(* IEC 61131-3 sources: daoli-st-library/DL_Process (part 23) *)

(* ---- FB_DL_BoilerThreeElement.st ---- *)
//==============================================================================
// 功能块：FB_DL_BoilerThreeElement ｜ 中文名称：锅炉三冲量给水控制（复杂度 H）
// 所属子库：DL_Process ｜ 版本：v1.0.0 ｜ 兼容：CODESYS V3.5+ / TwinCAT 3 / 汇川 InoProShop
// 功能描述：锅炉三冲量给水——汽包水位主回路（组合调用 FB_DL_PidController）
//           + 蒸汽流量前馈① + 给水流量反馈②，合成给水流量给定 [t/h]；
//           手/自无扰切换（跟踪）；蒸汽/给水流量比持续偏离判泄漏疑似。
// 开源溯源 (Origin)：道莅原创实现（参考锅炉三冲量给水控制工程惯例 分类与参数域）
// 单位表：水位[%] / 流量[t/h] / 增益[（t/h）/（t/h）] / 给定满量程[t/h] /
//         PID 参数[s] / 确认窗[ms] / 比偏阈[倍]
// 错误码表：16#0005_01EC 信息级（给水/蒸汽流量比持续超偏，泄漏疑似，
//           R13 三分类诊断范式，不置 bError）/ 16#0005_01ED 预留禁用
//           （不得挪用）/ 16#0005_0327 故障级（任一流量/水位非有限，保持
//           末次有效给定，切手动会扰动汽包，与 R22 CrossLimitSelect 同侧
//           策略，置 bError）/ 16#0005_0328 预留禁用（不得挪用）/
//           16#0005_0329 故障级兜底（置 bError）
// 状态机：N/A（手/自切换 + 前馈合成 + 比偏判窗为电平逻辑，无相位状态机）
// 边界行为：① 任一流量/水位非有限 → 保持末次有效给定 + 故障 0327（不
//           静默归零——切手动会扰动汽包）；② bAutoMode 下降沿 → 无扰切
//           手动（给定冻结为当前值）；③ 手动→自动无扰切换（PID 跟踪
//           注入当前给定）；④ 流量比超偏持续确认窗 → 信息 01EC；
//           ⑤ 给定下限钳 0（不倒转）；⑥ 非有限前馈增益 → 0327 复用。
// 依赖纪律：Process → Level 0/1 组合调用合法——水位主回路组合调用
//           FB_DL_PidController（DL_Algo，接口已核实：bEnable/bManual/
//           fSetpoint/fActual/fKp/tTi/tTd/rOutMin/rOutMax/bTrack/fTrackValue/
//           fOut），头注释依赖清单声明；蒸汽前馈律在本件内联（单乘法
//           合成属编排语义，非算法复制）。
// 修订历史：v1.0.0 2026-11-17 首版（R23 派单 · ROADMAP P1 §322）
//==============================================================================

FUNCTION_BLOCK FB_DL_BoilerThreeElement
VAR_INPUT
    fDrumLevelPct  : LREAL;                 // 汽包水位实测 [百分数] / Drum level [percent]
    fSteamFlowTh   : LREAL;                 // 蒸汽流量 [吨/小时]，前馈① / Steam flow [t/h], feedforward 1
    fFeedFlowTh    : LREAL;                 // 给水流量 [吨/小时]，反馈② / Feedwater flow [t/h], feedback 2
    fLevelSpPct    : LREAL := 50.0;         // 水位设定 [百分数] / Level setpoint [percent]
    fFwdGainSteam  : LREAL := 1.0;          // 蒸汽前馈增益 [（吨/小时）/（吨/小时）] / Steam feedforward gain
    fLevelKp       : LREAL := 2.0;          // 水位主回比例增益 [1] / Level loop proportional gain
    tLevelTi       : TIME  := T#30S;        // 水位主回积分时间 [s]，T#0S = 纯 PD / Level loop integral time [s]
    tLevelTd       : TIME  := T#0S;         // 水位主回微分时间 [s]，T#0S = 关闭 / Level loop derivative time [s]
    bAutoMode      : BOOL;                  // 自动模式请求 [—] / Auto mode request
    bReset         : BOOL;                  // 故障复位 [—] / Fault reset
END_VAR
VAR_OUTPUT
    fFeedSpTh      : LREAL;                 // 给水流量给定 [吨/小时] = PID 主回路 + 双前馈 / Feedwater setpoint [t/h] = PID plus feedforwards
    bAuto          : BOOL;                  // 实际自动态 [—] / Actual auto state
    eErr           : UDINT;                 // 错误码，0 = 无错 / Error code, 0 = no error
    bError         : BOOL;                  // 故障级标志，仅故障级错误置位 / Fault-class flag, set only on fault-level codes
    bValid         : BOOL;                  // 输出可用标志 / Outputs usable flag
END_VAR
VAR
    fbLevelPid     : FB_DL_PidController;   // 水位主回 PID（Level 0 组合调用） / Level loop PID, Level 0 composition
    fbRatioWin     : TON;                   // 流量比偏确认窗，段 6 无条件刷新 [ms] / Ratio-deviation confirm window
    _fFeedSpHeld   : LREAL;                 // 末次有效给定保持量 [吨/小时] / Held last valid setpoint [t/h]
    _fPidTrackPct  : LREAL;                 // 跟踪/手动值（PID % 域换算） [%] / Track and manual value in the PID percent domain
    _bAutoPrev     : BOOL;                  // 自动请求上拍电平快照 / Previous-scan auto request snapshot
    _bTrackNow     : BOOL;                  // 无扰投切跟踪当拍标志 / Bumpless track flag of this scan
    _bInit         : BOOL := FALSE;         // 首扫标志，初值 FALSE 取非判定 / First-scan flag, tested negated
    _bFiniteBad    : BOOL;                  // 非有限锁存 / Non-finite latch
    _bRatioSuspect : BOOL;                  // 比偏疑似当拍标志 / Ratio-suspect flag of this scan
    _bIllegal      : BOOL;                  // 非法状态标志 / Illegal state flag
END_VAR
VAR CONSTANT
    DL_BLR_SPAN_TH  : LREAL := 100.0;       // 给水给定满量程 [吨/小时]，PID 输出 [%] → [t/h] 映射基准 / Feedwater setpoint span [t/h], PID percent mapping base
    DL_BLR_RATIO_DEV: LREAL := 2.0;         // 给水/蒸汽比偏阈 [倍] / Feed-to-steam ratio deviation bound [ratio]
    DL_BLR_RATIO_WIN: TIME  := T#10S;       // 比偏确认窗 [ms] / Ratio-deviation confirm window [ms]
    DL_BLR_FLOW_MIN : LREAL := 1.0;         // 比偏判据流量下限 [吨/小时]，防小流量假比 / Ratio floor [t/h], guards a false ratio at low flows
    DL_BLR_INF      : LREAL := 1.7976931348623157E308; // LREAL 幅值上限 / LREAL magnitude ceiling
    DL_BLR_EPS      : LREAL := 1.0E-6;      // 浮点判零容差 / Float zero tolerance
END_VAR

(*------------------------------------------------------------------------------
 * 段 1｜每拍预置：给定保持量起步为零，单拍标志预清零
 *      Held setpoint starts at zero, one-shot flags pre-cleared
 *-----------------------------------------------------------------------------*)
fFeedSpTh := 0.0;                           // 给定预置零（异常路径由保持量覆盖） / Setpoint preset zero, held value overrides on anomaly
bAuto     := FALSE;                         // 自动态预置 FALSE / Auto preset FALSE
eErr      := 16#0000_0000;                  // 错误码每拍重算 / Error code recomputed
bError    := FALSE;                         // 故障标志每拍重算 / Fault flag recomputed
bValid    := FALSE;                         // 可用标志每拍重算 / Usable flag recomputed
_bTrackNow  := FALSE;                       // 跟踪标志预清零 / Track flag pre-cleared
_bRatioSuspect := FALSE;                    // 比偏标志预清零 / Ratio flag pre-cleared
_bIllegal   := FALSE;                       // 非法状态预清零 / Illegal flag pre-cleared

(*------------------------------------------------------------------------------
 * 段 2｜首扫初始化与手/自沿检测
 *      First-scan initialisation and the auto-edge detection
 *-----------------------------------------------------------------------------*)
IF NOT _bInit THEN
    _fFeedSpHeld := 0.0;                    // 保持量清零 / Held value cleared
    _bFiniteBad  := FALSE;                  // 非有限锁存清零 / Non-finite latch cleared
    _bInit       := TRUE;                   // 首扫只做一次 / The first scan runs once
END_IF
IF (NOT bAutoMode) AND _bAutoPrev THEN
    _bTrackNow := FALSE;                    // 下降沿：无扰切手动（给定冻结，PID bManual 承担） / Falling edge, bumpless to manual, the setpoint freezes
END_IF
IF bAutoMode AND (NOT _bAutoPrev) THEN
    _bTrackNow := TRUE;                     // 上升沿：无扰投切（PID 跟踪注入当前给定） / Rising edge, bumpless track injection
END_IF
_bAutoPrev := bAutoMode;                    // 电平快照推进 / Snapshot advanced

(*------------------------------------------------------------------------------
 * 段 3｜输入防御闸（任一流量/水位/增益非有限 → 0327，保持末值）
 *      Input defense gate, last held setpoint kept on anomaly
 *-----------------------------------------------------------------------------*)
IF (fDrumLevelPct <> fDrumLevelPct) OR (ABS(fDrumLevelPct) > DL_BLR_INF)
   OR (fSteamFlowTh <> fSteamFlowTh) OR (ABS(fSteamFlowTh) > DL_BLR_INF)
   OR (fFeedFlowTh <> fFeedFlowTh) OR (ABS(fFeedFlowTh) > DL_BLR_INF)
   OR (fLevelSpPct <> fLevelSpPct) OR (ABS(fLevelSpPct) > DL_BLR_INF)
   OR (fFwdGainSteam <> fFwdGainSteam) OR (ABS(fFwdGainSteam) > DL_BLR_INF) THEN
    _bFiniteBad := TRUE;                    // 非有限锁存 / Non-finite latched
END_IF
IF bReset THEN
    _bFiniteBad := FALSE;                   // 复位清非有限锁存 / Reset clears the latch
END_IF

(*------------------------------------------------------------------------------
 * 段 4｜PID 主回路组合调用（无条件周期刷新，R40：每拍必调）
 *      PID composition called unconditionally every scan per R40
 *-----------------------------------------------------------------------------*)
IF ABS(fFwdGainSteam) > DL_BLR_EPS THEN
    _fPidTrackPct := ((_fFeedSpHeld - fFwdGainSteam * fSteamFlowTh) / DL_BLR_SPAN_TH) * 100.0; // 当前给定反算 PID % 域跟踪值 / Current setpoint back-computed to the PID percent domain
ELSE
    _fPidTrackPct := (_fFeedSpHeld / DL_BLR_SPAN_TH) * 100.0; // 前馈增益为零：按纯主回换算 / Zero gain, pure loop conversion
END_IF
IF _fPidTrackPct < 0.0 THEN
    _fPidTrackPct := 0.0;                   // 跟踪值下限钳 0 / Track value lower clamp
ELSIF _fPidTrackPct > 100.0 THEN
    _fPidTrackPct := 100.0;                 // 跟踪值上限钳 100 / Track value ceiling clamp
END_IF
fbLevelPid(bEnable      := bAutoMode AND (NOT _bFiniteBad),
           bManual      := (NOT bAutoMode) OR _bFiniteBad,
           fManualValue := _fPidTrackPct,
           fSetpoint    := fLevelSpPct,
           fActual      := fDrumLevelPct,
           fKp          := fLevelKp,
           tTi          := tLevelTi,
           tTd          := tLevelTd,
           fDeadband    := 0.0,
           bIncremental := FALSE,
           rOutMin      := 0.0,
           rOutMax      := 100.0,
           bTrack       := _bTrackNow,
           fTrackValue  := _fPidTrackPct,
           bReset       := FALSE);         // 水位主回 PID / Level loop PID
IF _bTrackNow THEN
    _bTrackNow := FALSE;                    // 跟踪只注一拍（无扰投切窗口收敛） / Track injected for one scan only
END_IF

(*------------------------------------------------------------------------------
 * 段 5｜三冲量合成：给定 = PID 主回路换算 + 蒸汽前馈（内联合成）
 *      Three-element synthesis, feedforward inlined
 *-----------------------------------------------------------------------------*)
IF (NOT _bFiniteBad) THEN
    fFeedSpTh := (fbLevelPid.fOut / 100.0) * DL_BLR_SPAN_TH + fFwdGainSteam * fSteamFlowTh; // 三冲量给定 [吨/小时] / Three-element setpoint [t/h]
    IF fFeedSpTh < 0.0 THEN
        fFeedSpTh := 0.0;                   // 给定下限钳 0（不倒转） / Lower clamp, no reverse
    END_IF
    _fFeedSpHeld := fFeedSpTh;              // 末次有效给定保持量推进 / Held setpoint advanced
ELSE
    fFeedSpTh := _fFeedSpHeld;              // 异常路径：保持末次有效给定（0327 口径） / Anomaly, last held setpoint kept
END_IF
bAuto := bAutoMode AND (NOT _bFiniteBad);   // 实际自动态出口 / Actual auto outlet

(*------------------------------------------------------------------------------
 * 段 6｜流量比偏确认窗无条件刷新（R40：CASE 之外每拍必调）
 *      Ratio-deviation window refreshed unconditionally per R40
 *-----------------------------------------------------------------------------*)
IF (ABS(fSteamFlowTh) > DL_BLR_FLOW_MIN) AND (ABS(fFeedFlowTh) > DL_BLR_FLOW_MIN) THEN
    IF (fFeedFlowTh > fSteamFlowTh * DL_BLR_RATIO_DEV)
       OR (fSteamFlowTh > fFeedFlowTh * DL_BLR_RATIO_DEV) THEN
        _bRatioSuspect := TRUE;             // 双侧直比（禁 ABS 单侧，R19 整数纪律同源） / Two-sided direct comparison
    END_IF
END_IF
fbRatioWin(IN := bAutoMode AND (NOT _bFiniteBad) AND _bRatioSuspect, PT := DL_BLR_RATIO_WIN); // 比偏确认窗 / Ratio-deviation window

(*------------------------------------------------------------------------------
 * 段 7｜码位出口
 *      Code outlet
 *-----------------------------------------------------------------------------*)
IF _bIllegal THEN
    eErr   := 16#0005_0329;                 // 故障级：兜底 / Fault: fallback
    bError := TRUE;                         // 置故障标志 / Raise the fault flag
ELSIF _bFiniteBad THEN
    eErr   := 16#0005_0327;                 // 故障级：非有限输入保持末值 / Fault: non-finite input, held setpoint
    bError := TRUE;                         // 置故障标志（R45 配对） / Raise the fault flag
    bValid := FALSE;                        // 输出不可用 / Outputs unusable
ELSIF fbRatioWin.Q THEN
    eErr := 16#0005_01EC;                   // 信息级：流量比超偏，泄漏疑似 / Info: ratio deviation, leak suspected
    bValid := TRUE;                         // 输出可用 / Outputs usable
ELSE
    bValid := bAutoMode;                    // 自动态输出可用；手动态给定由调用方使用 / Usable in auto, the manual setpoint is for the caller
END_IF
END_FUNCTION_BLOCK

(* ---- FB_DL_BrewFermentTempRampSeq.st ---- *)
// FB_DL_BrewFermentTempRampSeq v1.0.0
// 开源溯源：clean-room 自研（族 DL_Process，ST 生态实测 0 命中，无外部代码引入）
(*
  功能: 发酵温度阶梯七相顺控：IDLE→PITCH→MAIN→REST→COOL→HOLD→IDLE 置 xDone。
        判据：PITCH 达 fPitchTemp±0.5 °C；MAIN 当 fExtract ≤ fExtractEnd；REST 满 48 h；
        COOL 达 fCoolTemp±0.5 °C；HOLD 满 24 h。设定值 _fSp 按 fRampRate [°C/h] 逐周期逼近目标，
        单周期增量 = fRampRate·fCycleS/3600 [°C]，严禁阶跃（相切换不回跳）。
        阀位：实测高于设定 0.2 °C 开冷却阀，低于 0.2 °C 开加热阀，两阀互斥，互锁复核失败双阀 FALSE 并锁存。
  邻件: 与 FC_DL_FermentAttenuationCalc、FC_DL_DiacetylRestWindowCalc、FC_DL_BeerCoolingLoadCalc 同族，本件不调用 FC。
  码表: 9341 入参非有限｜9342 组态非法(fRampRate/fCycleS≤0)｜9343 相超时(12/240/24 h)
        9344 温控失效或双阀互锁违例｜9345 相位落 ELSE 兜底｜9346 信息级序列完成。故障码锁存至 xReset 上升沿。
  边界: 无方法块/无属性块/无全局变量/无物理 IO 地址；六 TON 无条件刷新；温度非有限 → FAULT 且双阀 FALSE。
*)
TYPE E_DL_FermentRampPhase :
(
    IDLE  := 0,         // 空闲：等启动指令 [-] / Idle, waiting start
    PITCH := 10,        // 接种：控温至接种温度 [-] / Pitching temperature
    MAIN  := 20,        // 主发酵：控温至主发酵温度 [-] / Main fermentation
    REST  := 30,        // 还原：升温双乙酰还原 [-] / Diacetyl rest
    COOL  := 40,        // 降温：降至贮酒温度 [-] / Cooling down
    HOLD  := 50,        // 贮酒：低温保持 [-] / Cold holding
    FAULT := 90         // 故障：锁存，仅复位沿可出 [-] / Fault latched
);
END_TYPE
FUNCTION_BLOCK FB_DL_BrewFermentTempRampSeq
VAR_INPUT
    xEnable     : BOOL := FALSE;    // 使能，FALSE 时冻结在 IDLE [-] / Enable gate
    xStart      : BOOL := FALSE;    // 启动指令，上升沿有效 [-] / Start rising edge
    xReset      : BOOL := FALSE;    // 复位，上升沿清故障锁存 [-] / Reset rising edge
    fTankTemp   : REAL := 8.0;      // 罐内实测温度 [°C] / Measured tank temperature [degC]
    fPitchTemp  : REAL := 9.0;      // 接种温度设定 [°C] / Pitching temperature [degC]
    fMainTemp   : REAL := 11.0;     // 主发酵温度设定 [°C] / Main temperature [degC]
    fRestTemp   : REAL := 16.0;     // 还原温度设定 [°C] / Rest temperature [degC]
    fCoolTemp   : REAL := 1.0;      // 贮酒温度设定 [°C] / Cold storage temperature [degC]
    fRampRate   : REAL := 0.5;      // 斜坡速率 [°C/h]，域 > 0 / Ramp rate [degC/h]
    fExtract    : REAL := 12.0;     // 当前外观浓度 [°P] / Current extract [degP]
    fExtractEnd : REAL := 3.0;      // 主发酵终点浓度 [°P] / End-of-main extract [degP]
    fCycleS     : REAL := 0.01;     // 任务周期 [s]，域 > 0 / Task cycle time [s]
END_VAR
VAR_OUTPUT
    ePhase     : E_DL_FermentRampPhase;     // 相位出口，段尾单点映射 [-] / Phase outlet
    fTempSp    : REAL;                      // 温度设定出口 [°C] / Temperature setpoint outlet [degC]
    xCoolValve : BOOL;                      // 冷却阀指令 [-] / Cooling valve command
    xHeatValve : BOOL;                      // 加热阀指令 [-] / Heating valve command
    xDone      : BOOL;                      // 序列完成单拍脉冲 [-] / Done one-shot pulse
    xFault     : BOOL;                      // 故障锁存标志 [-] / Fault latch flag
    uErrorId   : UDINT;                     // 事件码，0 = 无事件 / Event code
END_VAR
VAR
    tonPitch  : TON;                        // 接种相超时 12 h，无条件刷新 / Pitch timeout
    tonMain   : TON;                        // 主发酵相超时 240 h，无条件刷新 / Main timeout
    tonRest   : TON;                        // 还原相定时 48 h，无条件刷新 / Rest timer
    tonCool   : TON;                        // 降温相超时 24 h，无条件刷新 / Cool timeout
    tonHold   : TON;                        // 贮酒相定时 24 h，无条件刷新 / Hold timer
    tonDev    : TON;                        // 温控偏差持续窗 600 s，无条件刷新 / Deviation window
    rtStart   : R_TRIG;                     // 启动沿实例，无条件刷新 / Start edge instance
    rtReset   : R_TRIG;                     // 复位沿实例，无条件刷新 / Reset edge instance
    _ePhase   : E_DL_FermentRampPhase := E_DL_FermentRampPhase.IDLE;    // 内部相位，CASE 唯一写入 / Internal phase
    _fSp      : REAL := 0.0;                // 温度设定斜坡量 [°C] / Ramp setpoint [degC]
    _fSpTar   : REAL := 0.0;                // 本相设定目标 [°C] / Phase setpoint target [degC]
    _fStep    : REAL := 0.0;                // 本周期斜坡增量 [°C] / Per-cycle ramp step [degC]
    _xCoolOn  : BOOL := FALSE;              // 冷却阀内部选择位 [-] / Internal cooling selection
    _xHeatOn  : BOOL := FALSE;              // 加热阀内部选择位 [-] / Internal heating selection
    _bFault   : BOOL := FALSE;              // 故障锁存位（锁存量，仅复位沿清）/ Latched fault bit
    _uFault   : UDINT := 16#0000;           // 故障码锁存（锁存量，仅复位沿清）/ Latched fault code
    _uInfo    : UDINT := 16#0000;           // 信息码，每拍重算 / Transient info code
END_VAR
// 段 0：定时器与沿实例无条件周期刷新（禁置于 IF/CASE 内，R7/R188）/ Unconditional refresh
rtStart(CLK := xStart);                                                     // 启动沿每拍必调 / Start edge
rtReset(CLK := xReset);                                                     // 复位沿每拍必调 / Reset edge
tonPitch(IN := (_ePhase = E_DL_FermentRampPhase.PITCH), PT := T#12H);       // 接种相超时 / Pitch timeout
tonMain(IN := (_ePhase = E_DL_FermentRampPhase.MAIN), PT := T#240H);        // 主发酵超时 / Main timeout
tonRest(IN := (_ePhase = E_DL_FermentRampPhase.REST), PT := T#48H);         // 还原 48 h / Rest timer
tonCool(IN := (_ePhase = E_DL_FermentRampPhase.COOL), PT := T#24H);         // 降温超时 / Cool timeout
tonHold(IN := (_ePhase = E_DL_FermentRampPhase.HOLD), PT := T#24H);         // 贮酒 24 h / Hold timer
tonDev(IN := (_ePhase <> E_DL_FermentRampPhase.IDLE) AND (_ePhase <> E_DL_FermentRampPhase.FAULT)
             AND (ABS(fTankTemp - _fSp) > 3.0), PT := T#600S);              // 温控偏差窗 / Deviation window
// 段 1：单拍量与阀位预清零（锁存量 _bFault/_uFault/_fSp 不入清单，R187）/ One-shot clear
_uInfo := 16#0000;                  // 信息码每拍重算 / Info code recomputed
xDone := FALSE;                     // 完成脉冲缺省清 / Done pulse clear
_xCoolOn := FALSE;                  // 冷却阀缺省关（互锁起点）/ Cooling default off
_xHeatOn := FALSE;                  // 加热阀缺省关（互锁起点）/ Heating default off
// 段 2：非有限闸与组态域闸（归因唯一，逐因独立码，R190）/ Gate stage
IF (fTankTemp <> fTankTemp) OR (fPitchTemp <> fPitchTemp) OR (fMainTemp <> fMainTemp)
   OR (fRestTemp <> fRestTemp) OR (fCoolTemp <> fCoolTemp) OR (fRampRate <> fRampRate)
   OR (fExtract <> fExtract) OR (fExtractEnd <> fExtractEnd) OR (fCycleS <> fCycleS)
   OR (ABS(fTankTemp) >= 3.0E38) OR (ABS(fPitchTemp) >= 3.0E38) OR (ABS(fMainTemp) >= 3.0E38)
   OR (ABS(fRestTemp) >= 3.0E38) OR (ABS(fCoolTemp) >= 3.0E38) OR (ABS(fRampRate) >= 3.0E38)
   OR (ABS(fExtract) >= 3.0E38) OR (ABS(fExtractEnd) >= 3.0E38) OR (ABS(fCycleS) >= 3.0E38) THEN
    _uFault := 16#0002_9341;        // 故障级：入参非有限 / Fault: non-finite input
    _bFault := TRUE;                // 置故障锁存（R45 配对）/ Set fault latch
END_IF
IF (fRampRate <= 1.0E-9) OR (fCycleS <= 1.0E-6) THEN
    _uFault := 16#0002_9342;        // 故障级：组态非法 / Fault: illegal configuration
    _bFault := TRUE;                // 置故障锁存（R45 配对）/ Set fault latch
END_IF
// 段 3：温控失效持续窗（偏差超 3 °C 达 600 s）/ Control deviation window
IF tonDev.Q THEN
    _uFault := 16#0002_9344;        // 故障级：温控失效 / Fault: control failure
    _bFault := TRUE;                // 置故障锁存（R45 配对）/ Set fault latch
END_IF
// 段 4：复位沿（FAULT 唯一解除路径）/ Reset edge, only exit from fault
IF rtReset.Q THEN                   // rtReset.Q = 当拍量 / Reset edge per scan
    IF _ePhase = E_DL_FermentRampPhase.FAULT THEN
        _ePhase := E_DL_FermentRampPhase.IDLE;      // 故障相迁出回空闲 / Fault exits to idle
    END_IF
    _fSp := fTankTemp;              // 设定回实测（复位不阶跃）/ Setpoint resumes at measured value
    _bFault := FALSE;               // 清故障锁存位（仅此解除沿可清）/ Clear latched bit
    _uFault := 16#0000;             // 清故障锁存码（仅此解除沿可清）/ Clear latched code
END_IF
// 段 5：相位机（先消化本拍合法事件，再消化超时，R275）/ Phase machine
CASE _ePhase OF
E_DL_FermentRampPhase.IDLE:
    _fSp := fTankTemp;                              // 空闲设定随实测（无阶跃）/ Track measured value
    IF _bFault THEN
        _ePhase := E_DL_FermentRampPhase.FAULT;     // 聚合故障进故障相 / Enter fault
    ELSIF rtStart.Q AND xEnable THEN
        _ePhase := E_DL_FermentRampPhase.PITCH;     // 启动：进接种相 / Start, pitching
    END_IF
E_DL_FermentRampPhase.PITCH:
    _fSpTar := fPitchTemp;                          // 接种相目标 / Pitching target
    IF _bFault THEN
        _ePhase := E_DL_FermentRampPhase.FAULT;     // 故障优先 / Fault first
    ELSIF NOT xEnable THEN
        _ePhase := E_DL_FermentRampPhase.IDLE;      // 使能撤销回空闲 / Enable dropped
    ELSIF ABS(fTankTemp - fPitchTemp) <= 0.5 THEN
        _ePhase := E_DL_FermentRampPhase.MAIN;      // 达 ±0.5 °C：进主发酵相 / Go main
    ELSIF tonPitch.Q THEN
        _uFault := 16#0002_9343;                    // 故障级：接种相超时 / Pitch timeout
        _bFault := TRUE;                            // 置故障锁存（R45 配对）/ Set latch
        _ePhase := E_DL_FermentRampPhase.FAULT;     // 进故障相 / Enter fault
    END_IF
E_DL_FermentRampPhase.MAIN:
    _fSpTar := fMainTemp;                           // 主发酵目标 / Main target
    IF _bFault THEN
        _ePhase := E_DL_FermentRampPhase.FAULT;     // 故障优先 / Fault first
    ELSIF NOT xEnable THEN
        _ePhase := E_DL_FermentRampPhase.IDLE;      // 使能撤销回空闲 / Enable dropped
    ELSIF fExtract <= fExtractEnd THEN
        _ePhase := E_DL_FermentRampPhase.REST;      // 浓度达终点：进还原相 / Go rest
    ELSIF tonMain.Q THEN
        _uFault := 16#0002_9343;                    // 故障级：主发酵相超时 / Main timeout
        _bFault := TRUE;                            // 置故障锁存（R45 配对）/ Set latch
        _ePhase := E_DL_FermentRampPhase.FAULT;     // 进故障相 / Enter fault
    END_IF
E_DL_FermentRampPhase.REST:
    _fSpTar := fRestTemp;                           // 还原温度目标 / Rest target
    IF _bFault THEN
        _ePhase := E_DL_FermentRampPhase.FAULT;     // 故障优先 / Fault first
    ELSIF tonRest.Q THEN
        _ePhase := E_DL_FermentRampPhase.COOL;      // 满 48 h：进降温相 / Rest done, cool
    END_IF
E_DL_FermentRampPhase.COOL:
    _fSpTar := fCoolTemp;                           // 降温目标 / Cooling target
    IF _bFault THEN
        _ePhase := E_DL_FermentRampPhase.FAULT;     // 故障优先 / Fault first
    ELSIF ABS(fTankTemp - fCoolTemp) <= 0.5 THEN
        _ePhase := E_DL_FermentRampPhase.HOLD;      // 达贮酒温度：进贮酒相 / Go hold
    ELSIF tonCool.Q THEN
        _uFault := 16#0002_9343;                    // 故障级：降温相超时 / Cool timeout
        _bFault := TRUE;                            // 置故障锁存（R45 配对）/ Set latch
        _ePhase := E_DL_FermentRampPhase.FAULT;     // 进故障相 / Enter fault
    END_IF
E_DL_FermentRampPhase.HOLD:
    _fSpTar := fCoolTemp;                           // 贮酒温度保持 / Hold target
    IF _bFault THEN
        _ePhase := E_DL_FermentRampPhase.FAULT;     // 故障优先 / Fault first
    ELSIF tonHold.Q THEN
        xDone := TRUE;                              // 满 24 h：完成脉冲单拍 / Done pulse
        _uInfo := 16#0002_9346;                     // 信息级：序列完成 / Info: sequence done
        _ePhase := E_DL_FermentRampPhase.IDLE;      // 回空闲 / Return to idle
    END_IF
E_DL_FermentRampPhase.FAULT:
    _fSpTar := fTankTemp;                           // 故障相设定回实测 / Setpoint tracks measured
    IF rtReset.Q THEN
        _ePhase := E_DL_FermentRampPhase.IDLE;      // 复位沿解除（段 4 已清锁存）/ Reset releases
    END_IF
ELSE
    _uFault := 16#0002_9345;                        // 故障级：非法相位兜底 / Illegal phase id
    _bFault := TRUE;                                // 置故障锁存（R45 配对）/ Set latch
    _fSpTar := fTankTemp;                           // 非法相位设定回实测 / Setpoint tracks measured
    _ePhase := E_DL_FermentRampPhase.FAULT;         // 强制进故障相 / Force into fault
END_CASE
// 段 6：设定值斜坡（增量 = fRampRate·fCycleS/3600，禁阶跃）/ Setpoint ramp
IF (_ePhase = E_DL_FermentRampPhase.IDLE) OR (_ePhase = E_DL_FermentRampPhase.FAULT) THEN
    _fSp := fTankTemp;                              // 空闲/故障相跟随实测 / Track measured value
ELSE
    _fStep := fRampRate * fCycleS / 3600.0;         // 本周期增量 [°C] / Per-cycle step
    IF _fSp < _fSpTar THEN
        _fSp := _fSp + _fStep;                      // 向上逼近 / Ramp upward
        IF _fSp > _fSpTar THEN
            _fSp := _fSpTar;                        // 不得越过目标 / No overshoot
        END_IF
    ELSIF _fSp > _fSpTar THEN
        _fSp := _fSp - _fStep;                      // 向下逼近 / Ramp downward
        IF _fSp < _fSpTar THEN
            _fSp := _fSpTar;                        // 不得越过目标 / No overshoot
        END_IF
    END_IF
END_IF
// 段 7：阀位生成（实测高于设定 0.2 °C 开冷阀，反之开热阀，互斥）/ Valve generation
IF (_ePhase = E_DL_FermentRampPhase.IDLE) OR (_ePhase = E_DL_FermentRampPhase.FAULT) THEN
    _xCoolOn := FALSE;                              // 空闲/故障相不推阀 / No valve action
    _xHeatOn := FALSE;                              // 空闲/故障相不推阀 / No valve action
ELSIF (fTankTemp - _fSp) > 0.2 THEN
    _xCoolOn := TRUE;                               // 偏热：开冷却阀 / Too warm, cool
ELSIF (fTankTemp - _fSp) < -0.2 THEN
    _xHeatOn := TRUE;                               // 偏冷：开加热阀 / Too cold, heat
END_IF
// 段 8：出口单点映射（名实双出口，R191；双阀互锁复核）/ Outlet mapping
ePhase := _ePhase;                                  // 相位出口单点映射 / Phase outlet
IF (_ePhase = E_DL_FermentRampPhase.FAULT) OR _bFault THEN
    fTempSp := fTankTemp;                           // 故障侧设定跟随实测 / Setpoint tracks measured
    xCoolValve := FALSE;                            // 故障侧冷却阀硬关 / Cooling hard off
    xHeatValve := FALSE;                            // 故障侧加热阀硬关 / Heating hard off
    xFault := TRUE;                                 // 故障锁存回放 / Replay latched flag
    uErrorId := _uFault;                            // 故障码锁存回放 / Replay latched code
ELSIF _xCoolOn AND _xHeatOn THEN
    fTempSp := _fSp;                                // 设定值出口 / Setpoint outlet
    xCoolValve := FALSE;                            // 互锁违例：双阀全关 / Interlock: both off
    xHeatValve := FALSE;                            // 互锁违例：双阀全关 / Interlock: both off
    xFault := TRUE;                                 // 互锁违例置故障 / Raise fault on interlock
    uErrorId := 16#0002_9344;                       // 故障级：双阀互锁违例 / Fault: valve interlock
ELSE
    fTempSp := _fSp;                                // 设定值出口 / Setpoint outlet
    xCoolValve := _xCoolOn;                         // 冷却阀出口 / Cooling outlet
    xHeatValve := _xHeatOn;                         // 加热阀出口 / Heating outlet
    xFault := FALSE;                                // 无故障 / No fault
    uErrorId := _uInfo;                             // 信息码每拍重算 / Transient info code
END_IF
IF (fTempSp <> fTempSp) OR (ABS(fTempSp) >= 3.0E38) THEN
    fTempSp := fTankTemp;                           // 出口复核失败回实测 / Outlet recheck fallback
    xCoolValve := FALSE;                            // 出口复核失败关冷却 / Cut cooling
    xHeatValve := FALSE;                            // 出口复核失败关加热 / Cut heating
    xFault := TRUE;                                 // 出口复核失败置故障 / Raise fault
    uErrorId := 16#0002_9341;                       // 故障级：出口非有限 / Fault: non-finite outlet
END_IF
END_FUNCTION_BLOCK

(* ---- FB_DL_BundleShrinkTemp.st ---- *)
(*
  FB_DL_BundleShrinkTemp  —  收缩包装热风温度窗（超温/欠温双判 + 冷却延时） / Shrink-wrap hot-air temperature window with over/under-temperature judgement and cooling delay
  分类 Category : DL_Process
  版本 Version  : 1.0.0
  来源 Source   : roadmap-pkg-p2 — 后道收缩包装工站真缺口
  溯源 Origin   : 道莅 clean-room 实现；热风升温-恒温-冷却三段与温度窗双判为公开包装工艺逻辑，未复制任何源码行
  功能 Function : 1) 三段顺控：eHeat 加热（温度进窗 [fTempLoC, fTempHiC] 后由 tHeat 计时，
                  升温超时视为欠温故障）→ eCool 冷却（tCool 到时）→ eDone；
                  2) 超温/欠温双判独立归因（eOverTemp / eUnderTemp，R190 禁共用成员）；
                  3) 故障级单码 03A5，归因由 eCause 独立成员承载；
                  4) 信息级 04CD = 收缩循环完成沿；5) 解除式全当拍量（R240）。
  接口 Interface: 输入热风温度/温度窗/升温与冷却时间；输出状态 + 窗内镜像 + 码
  边界 Boundary : ① 组态闸：fTempHiC <= fTempLoC、tHeat <= T#0S、tCool <= T#0S → 03A5 锁存；
                  ② 温度判据为双向容差式（下限 -1.0E-6 / 上限 +1.0E-6），禁 = / <> 判等；
                  ③ 升温超时仅在温度未进窗时成立（门控为相量而非单拍标志，禁 bError 门控）；
                  ④ 两个 TON + 一个 R_TRIG 段 0 无条件周期调用，IN 由相位派生；
                  ⑤ 故障相迁出唯一路径 = bReset 上升沿；⑥ 零全局耦合（无 GVL / %I %Q %M）。
  依赖 Depends  : Standard.library（TON / R_TRIG）
  码表 Error codes（Process 段 0005，故障窗口 03A5 / 信息窗口 04CD）:
    16#0005_03A5 故障级：收缩包装温度故障总码（组态非法 / 超温 / 欠温或升温超时），
                 锁存至 bReset 上升沿；归因见 eCause，不新增码位（派单硬约束单码）
    16#0005_04CD 信息级：收缩循环完成沿（冷却完成进 eDone 单拍）
  修订历史 Revision :
    2026-11-19  v1.0.0  R43 首版（批次 2 · 序号 9）
*)

TYPE E_DL_BstState :
(
    eIdle  := 0,      // 未使能待启动 / Idle, waiting start
    eHeat  := 10,     // 加热（温度窗 + 恒温计时） / Heating under window and dwell timing
    eCool  := 20,     // 冷却延时 / Cooling delay
    eDone  := 50,     // 循环完成 / Done
    eFault := 90      // 故障锁存相（加热输出冻结关断） / Fault latched, heater frozen off
);
END_TYPE

TYPE E_DL_BstCause :
(
    eNone       := 0, // 无故障成因 / No cause
    eCfgIllegal := 1, // 组态非法 / Illegal configuration
    eOverTemp   := 2, // 超温 / Over temperature
    eUnderTemp  := 3  // 欠温（含升温超时） / Under temperature including heat timeout
);
END_TYPE

FUNCTION_BLOCK FB_DL_BundleShrinkTemp
VAR_INPUT
    fTempC     : REAL := 0.0;         // 热风实测温度 [°C] / Measured hot-air temperature
    fTempLoC   : REAL := 150.0;       // 温度窗下限 [°C] / Temperature window low
    fTempHiC   : REAL := 180.0;       // 温度窗上限 [°C] / Temperature window high
    tHeat      : TIME := T#6S;        // 恒温保持时长 [ms]，域 > 0 / Heat dwell duration
    tCool      : TIME := T#3S;        // 冷却延时 [ms]，域 > 0 / Cooling delay
    bHeaterOn  : BOOL := FALSE;       // 加热使能（电平）[-] / Heater enable
    bStart     : BOOL := FALSE;       // 启动命令（电平）[-] / Start command
    bReset     : BOOL := FALSE;       // 复位命令，上升沿清故障 [-] / Reset edge
END_VAR
VAR_OUTPUT
    eState     : E_DL_BstState;       // 状态出口，段 6 单点映射 / State outlet
    eCause     : E_DL_BstCause;       // 故障成因出口（R190） / Fault cause outlet
    bHeaterCmd : BOOL;                // 加热输出指令 [-] / Heater command
    bInWindow  : BOOL;                // 温度在窗镜像 [-] / In-window mirror
    bCycleDone : BOOL;                // 循环完成标志 [-] / Cycle done flag
    bError     : BOOL;                // 故障锁存标志 [-] / Fault latch flag
    nErrId     : UDINT;               // 事件码，0 = 无事件 / Event code
END_VAR
VAR
    _eState    : E_DL_BstState := E_DL_BstState.eIdle;   // 内部相位（CASE 唯一写入目标） / Internal phase
    _eCause    : E_DL_BstCause := E_DL_BstCause.eNone;   // 故障成因锁存（锁存量） / Latched cause
    tonHeat    : TON;                 // 恒温保持计时，每周期无条件调用 / Heat dwell timer
    tonCool    : TON;                 // 冷却延时计时，每周期无条件调用 / Cooling timer
    rtReset    : R_TRIG;              // 复位沿实例，每周期无条件调用 / Reset edge
    _bWinOk    : BOOL;                // 温度在窗当拍量 [-] / In-window verdict
    _bOver     : BOOL;                // 超温当拍量 [-] / Over-temperature verdict
    _bCfgBad   : BOOL;                // 组态非法当拍量 [-] / Config illegal
    _bFault    : BOOL;                // 故障锁存位（锁存量） / Latched fault bit
    _uFault    : UDINT;               // 故障码锁存（锁存量） / Latched fault code
    _uInfo     : UDINT;               // 信息码，每拍重算 / Transient info code
END_VAR

(* —— 段 0：沿实例与定时器无条件周期刷新 + 当拍量判据 —— *)
_bWinOk := (fTempC >= fTempLoC - 1.0E-6) AND (fTempC <= fTempHiC + 1.0E-6);   // 温度容差窗判据 / Window verdict
_bOver := fTempC > (fTempHiC + 1.0E-6);                                      // 超温当拍量（上侧直比） / Over-temperature
_bCfgBad := (fTempHiC <= fTempLoC) OR (tHeat <= T#0S) OR (tCool <= T#0S);     // 组态非法当拍量 / Config illegal
rtReset(CLK := bReset);                                                      // 复位沿，每拍必调 / Reset edge
tonHeat(IN := (_eState = E_DL_BstState.eHeat), PT := tHeat);                 // 恒温保持计时 / Dwell timer
tonCool(IN := (_eState = E_DL_BstState.eCool), PT := tCool);                 // 冷却延时计时 / Cooling timer

(* —— 段 1：单拍量预清零（锁存量不入清单） —— *)
_uInfo := 16#0000_0000;            // 信息码每拍重算 / Info recomputed
bHeaterCmd := FALSE;               // 加热指令缺省关 / Heater command default off
bInWindow := FALSE;                // 窗内镜像缺省 FALSE / Window mirror default
bCycleDone := FALSE;               // 完成标志缺省 FALSE / Done default
nErrId := 16#0000_0000;            // 事件码缺省无事件 / Event code default

(* —— 段 2：复位沿 + 组态域闸 —— *)
IF rtReset.Q THEN                              // rtReset.Q = 当拍量 / current scan
    _bFault := FALSE;                          // 清故障锁存位（锁存量） / Clear fault latch
    _uFault := 16#0000_0000;                   // 清故障锁存码（锁存量） / Clear fault code
    _eCause := E_DL_BstCause.eNone;            // 清成因（锁存量） / Clear cause
    IF _eState = E_DL_BstState.eFault THEN
        _eState := E_DL_BstState.eIdle;        // 故障相迁出：回未使能 / Fault exit to idle
    END_IF
END_IF
IF _bCfgBad THEN                               // 组态域闸 / Config gate
    _uFault := 16#0005_03A5;                   // 故障级：温度故障总码 / Process fault code
    _eCause := E_DL_BstCause.eCfgIllegal;      // 归因：组态非法 / Cause: illegal config
    _bFault := TRUE;                           // 标志与码位配对（R45） / Flag paired with code
END_IF

(* —— 段 3：超温 / 欠温 / 升温超时（判据当拍量，门控为相位量） —— *)
IF (NOT _bFault) AND (_eState = E_DL_BstState.eHeat) AND _bOver THEN   // 超温 / Over temperature
    _uFault := 16#0005_03A5;
    _eCause := E_DL_BstCause.eOverTemp;        // 归因：超温 / Cause: over temperature
    _bFault := TRUE;
END_IF
IF (NOT _bFault) AND (_eState = E_DL_BstState.eHeat) AND (NOT _bWinOk) AND (NOT tonHeat.Q)
   AND (fTempC < (fTempLoC - 1.0E-6)) THEN     // 欠温（低于下限且计时未完成） / Under temperature
    _uFault := 16#0005_03A5;
    _eCause := E_DL_BstCause.eUnderTemp;       // 归因：欠温 / Cause: under temperature
    _bFault := TRUE;
END_IF
IF (NOT _bFault) AND (_eState = E_DL_BstState.eHeat) AND (NOT _bWinOk) AND tonHeat.Q THEN
    _uFault := 16#0005_03A5;
    _eCause := E_DL_BstCause.eUnderTemp;       // 归因：升温超时归并欠温 / Cause: heat timeout as under temp
    _bFault := TRUE;
END_IF

(* —— 段 4：故障解除式（R240；全当拍量）：rtReset.Q / NOT _bCfgBad / NOT _bOver / NOT _bWinOk 的当拍态 —— *)
IF rtReset.Q AND (NOT _bCfgBad) AND (NOT _bOver) THEN
    _bFault := FALSE;                          // 清故障锁存位（锁存量） / Clear fault latch
    _uFault := 16#0000_0000;                   // 清故障锁存码（锁存量） / Clear fault code
    _eCause := E_DL_BstCause.eNone;            // 清成因（锁存量） / Clear cause
END_IF

(* —— 段 4A：故障锁存相位迁移闸 —— *)
IF _bFault AND (_eState <> E_DL_BstState.eFault) THEN
    _eState := E_DL_BstState.eFault;           // 锁存即入故障相（加热关断） / Latch enters fault phase
END_IF

(* —— 段 5：相位机（CASE 全覆盖 + ELSE 兜底） —— *)
CASE _eState OF

E_DL_BstState.eIdle:
    IF bStart AND bHeaterOn AND (NOT _bFault) THEN   // 启动条件（须加热使能） / Start gate
        _eState := E_DL_BstState.eHeat;              // 进加热相 / Enter heating
    END_IF

E_DL_BstState.eHeat:
    bHeaterCmd := bHeaterOn;                         // 加热指令跟随使能（相内承载） / Heater command in phase
    IF tonHeat.Q AND _bWinOk THEN                    // 出口 1：恒温到时且在窗 / Dwell done in window
        _eState := E_DL_BstState.eCool;              // 进冷却相 / Enter cooling
    ELSIF (NOT bStart) OR (NOT bHeaterOn) THEN       // 出口 2：撤启动或撤加热（R98 双出口） / Start or heater released
        _eState := E_DL_BstState.eIdle;
    END_IF

E_DL_BstState.eCool:
    IF tonCool.Q THEN                                // 冷却到时 / Cooling elapsed
        _uInfo := 16#0005_04CD;                      // 信息级：收缩循环完成沿 / Info: cycle complete
        _eState := E_DL_BstState.eDone;              // 进完成相 / Enter done
    ELSIF NOT bStart THEN                            // 撤启动：中止 / Abort
        _eState := E_DL_BstState.eIdle;
    END_IF

E_DL_BstState.eDone:
    IF NOT bStart THEN                               // 撤启动回空闲 / Start released returns idle
        _eState := E_DL_BstState.eIdle;
    END_IF

E_DL_BstState.eFault:
    ;                                                // 故障相：加热关断，仅段 4 复位沿可迁出 / Heater off, reset only

ELSE
    _uFault := 16#0005_03A5;                   // 故障级：非法相位兜底（归并总码） / Illegal phase fallback
    _eCause := E_DL_BstCause.eCfgIllegal;      // 归因：相位非法归并组态 / Cause: phase illegal
    _bFault := TRUE;
    _eState := E_DL_BstState.eFault;           // 强制回故障相 / Force fault phase

END_CASE

(* —— 段 6：出口单点映射（名实同源；故障相加热强制关断） —— *)
IF _bFault THEN
    bHeaterCmd := FALSE;                       // 故障相加热强制关断（安全侧） / Heater forced off
    nErrId := _uFault;                         // 故障锁存码回放 / Replay latched code
ELSE
    nErrId := _uInfo;                          // 信息码 / Transient info
END_IF
bInWindow := _bWinOk AND (NOT _bFault);        // 窗内镜像 / Window mirror
bCycleDone := (_eState = E_DL_BstState.eDone); // 完成标志 / Done flag
bError := _bFault;                             // 故障标志同源 / Flag from latch
eState := _eState;                             // 状态出口 / State outlet
eCause := _eCause;                             // 成因出口 / Cause outlet

END_FUNCTION_BLOCK

(* ---- FB_DL_BusbarWeldMonitor.st ---- *)
(*==============================================================================
 * 组件名称 (Component)  : FB_DL_BusbarWeldMonitor
 * 所属子库 (Sublibrary) : DL_Process
 * 归属目录 (Directory)  : C:\Library\DL_Process
 * 当前版本 (Version)    : 1.0.0
 * 分类/来源标签         : 功能块（FUNCTION_BLOCK）· 母线焊接 · 超声焊能量包络
 *                         industry-pool / pvbusbar / ultrasonic-weld / envelope
 * 兼容性   (Platform)   : CODESYS 3.5 / TwinCAT 3 / 汇川 InoProShop / 施耐德
 *                         Machine Expert；仅用 Standard.library 的 TON / F_TRIG / ABS
 * 溯源声明 (Provenance) : 道莅自研 clean-room——只借公开规范条款与工程惯例，零代码行复制。
 * 功能一句话 (Summary)  : Busbar 超声焊接三维能量包络监视（功率-振幅-时间），
 *                         焊接期间任一维越窗即记缺陷，焊毕按在窗占比判定。
 *
 * 功能描述 (Function)   : 焊接进行中每拍评估三维窗口（功率带、振幅带、焊接
 *                         时长上限），任一维越窗当拍即置缺陷标记；焊接结束
 *                         （F_TRIG 下降沿）按在窗拍占比判定合格（信息级）或
 *                         缺陷（故障级）；时长越上限强制判缺陷并锁存；输入
 *                         非有限冻结监视。判定锁存到下一焊次起动沿解除。
 * 与既有件边界 (Boundary): 与库内激光焊轨迹件 LaserTabWeldTrack 为不同物理
 *                         域不同机制；本件只做包络判定，不出焊接功率给定。
 * 码位说明 (Codes)      : 信息 16#0006_3032 焊接判定合格（在窗占比达标）
 *                         故障 16#0006_3033 焊接判定缺陷（在窗占比不足）
 *                         故障 16#0006_3034 焊接时长越上限，强制缺陷
 *                         故障 16#0006_3035 输入非有限，监视冻结
 *                         段 16#06_0_32~36 首槽信息级、次槽起故障级。
 * 依赖说明 (Depends)    : 无 DL_ 内部依赖；仅 Standard.library 的 TON / F_TRIG。
 * 红线自检 (Redline)    : 零全局依赖 ｜ 零 VAR_EXTERNAL ｜ 零 %I/%Q ｜ 纯 IEC 标准库
 *                         NaN/Inf 精确判据拦截 ｜ 浮点比较带 fEps 容差
 *                         ENUM 配 CASE 且 ELSE 兜底 ｜ TON/F_TRIG 每周期无条件刷新
 *                         全变量双语同行注释 ｜ 判定锁存回放且有可达解除路径
 * 修订历史 (Revision)   : 2026-11-18  v1.0.0  首版入库（R32 · 批 4）
 *============================================================================*)

FUNCTION_BLOCK FB_DL_BusbarWeldMonitor
VAR_INPUT
    bRun     : BOOL;                    // 监视使能 / Enable
    bWelding : BOOL;                    // 焊接进行中 [事件] / Welding in progress
    fPowerKw : LREAL;                   // 焊接功率 [kW] / Welding power
    fAmpUm   : LREAL;                   // 振幅 [um] / Ultrasonic amplitude
    fPwrLoKw : LREAL := 4.0;            // 功率窗下限 [kW] / Power window lower bound
    fPwrHiKw : LREAL := 6.0;            // 功率窗上限 [kW] / Power window upper bound
    fAmpLoUm : LREAL := 35.0;           // 振幅窗下限 [um] / Amplitude window lower bound
    fAmpHiUm : LREAL := 55.0;           // 振幅窗上限 [um] / Amplitude window upper bound
    tWeldMaxS: TIME  := T#5S;           // 焊接时长上限 [s] / Weld duration limit
    fRatioTh : LREAL := 0.9;            // 在窗占比合格阈 [比值] / In-window ratio threshold
    fEps     : LREAL := 1.0E-6;         // 浮点判零容差 [实数域] / Floating zero tolerance
END_VAR
VAR_OUTPUT
    eVerdict : (ePending := 0, eGood := 1, eDefect := 2);       // 判定枚举输出 / Verdict output enum
    bInWin   : BOOL;                    // 当前拍三维都在窗内 / All three in window this scan
    fWinRatio: LREAL;                   // 在窗拍占比 [比值] / In-window scan ratio
    bError   : BOOL;                    // 故障标志，与故障码配对 / Fault flag paired with codes
    uErrorId : UDINT;                   // 事件码，0 表示无事件 / Event code, zero means none
END_VAR
VAR
    _eVerdict: (ePending := 0, eGood := 1, eDefect := 2);       // 内部判定 / Internal verdict
    tonWeld  : TON;     // 焊接时长计时 [s]，每拍无条件刷新 / Weld duration timer
    fTrigEnd : F_TRIG;  // 焊接结束下降沿，每拍无条件刷新 / Weld end falling edge
    bSigOk   : BOOL;    // 输入有效标志 / Input validity flag
    bWinNow  : BOOL;    // 本拍在窗判定 / This-scan window verdict
    nWinScans: UDINT;   // 在窗拍计数 [拍] / In-window scan count
    nTotScans: UDINT;   // 总拍计数 [拍] / Total scan count
    bTimeout : BOOL;    // 时长越限锁存 / Duration timeout latched
    bNewWeld : BOOL;    // 新焊次起动沿（焊接上升沿）/ New weld rising edge
    bPrevWld : BOOL;    // 上拍焊接快照 [开关] / Previous welding snapshot
    uCode    : UDINT;   // 码位暂存，出口单点写入 [码] / Code staging
END_VAR
VAR CONSTANT
    DL_BWM_PCT   : LREAL := 100.0;      // 百分比系数 [％] / Percent factor
    DL_BWM_BIGUD : UDINT := 4294967290; // 计数防回卷余量 [拍] / Counter wrap guard
END_VAR

(* 段 1｜定时器与边沿无条件刷新（红线 7）/ Timers and edges refreshed unconditionally *)
tonWeld(IN := bWelding AND bRun, PT := tWeldMaxS);  // 时长计时 / Duration timing
fTrigEnd(CLK := bWelding);                          // 焊接结束沿 / Weld end edge
bNewWeld := bWelding AND (NOT bPrevWld);            // 新焊次上升沿 / New weld edge
bPrevWld := bWelding;                               // 快照更新 / Update the snapshot

(* 段 2｜输入有效性（NaN 自反、Inf 上限）/ Input validity *)
bSigOk := (fPowerKw = fPowerKw) AND (fAmpUm = fAmpUm)               // NaN 自反判据 / NaN reflexivity
          AND (ABS(fPowerKw) < 1.0E308) AND (ABS(fAmpUm) < 1.0E308); // Inf 上限判据 / Inf limit

(* 段 3｜新焊次部署：计数清零，判定回待定，锁存解除（可达解除路径）
 *      New weld deployment: counters cleared, verdict reset, latch released *)
IF bNewWeld AND bRun THEN
    nWinScans := 0;                     // 在窗计数清零 / Clear the in-window count
    nTotScans := 0;                     // 总计数清零 / Clear the total count
    bTimeout := FALSE;                  // 时长锁存解除 / Release the timeout latch
    _eVerdict := ePending;              // 判定回待定 / Verdict to pending
    uCode := 16#0000_0000;              // 清码 / Clear the code
END_IF

(* 段 4｜焊接中每拍三维评估 / Per-scan three-dimension evaluation while welding *)
bWinNow := FALSE;                       // 默认不在窗 / Default out of window
IF bRun AND bWelding THEN
    IF NOT bSigOk THEN
        uCode := 16#0006_3035;          // 故障级：输入非有限，监视冻结 / Fault: frozen
    ELSE
        bWinNow := (fPowerKw >= fPwrLoKw - fEps) AND (fPowerKw <= fPwrHiKw + fEps)  // 功率在窗 / Power inside
                   AND (fAmpUm >= fAmpLoUm - fEps) AND (fAmpUm <= fAmpHiUm + fEps);  // 振幅在窗 / Amplitude inside
        nTotScans := nTotScans + 1;     // 总拍计数 / Count the scan
        IF bWinNow THEN
            nWinScans := nWinScans + 1; // 在窗计数 / Count in-window
        END_IF
        IF nTotScans >= DL_BWM_BIGUD THEN
            nTotScans := DL_BWM_BIGUD;  // 防回卷钳位 / Anti-wrap clamp
            nWinScans := nWinScans;     // 保持现值，占比保守 / Hold, ratio conservative
        END_IF
        IF tonWeld.Q THEN
            bTimeout := TRUE;           // 时长越限锁存 / Latch the timeout
        END_IF
    END_IF
END_IF
bInWin := bWinNow;                      // 在窗标志输出 / Window flag output

(* 段 5｜焊毕判定（F_TRIG 触发一次）：占比判合格或缺陷 / Verdict on weld end *)
IF fTrigEnd.Q AND bRun THEN
    IF (nTotScans > 0) AND (NOT bTimeout) THEN
        fWinRatio := UDINT_TO_LREAL(nWinScans) / UDINT_TO_LREAL(nTotScans);     // 占比导出 / Derive the ratio
        IF fWinRatio >= fRatioTh THEN
            _eVerdict := eGood;         // 判定合格 / Verdict good
            uCode := 16#0006_3032;      // 信息级：合格 / Info: good
        ELSE
            _eVerdict := eDefect;       // 判定缺陷 / Verdict defect
            uCode := 16#0006_3033;      // 故障级：占比不足 / Fault: ratio short
        END_IF
    ELSIF bTimeout THEN
        _eVerdict := eDefect;           // 超时强制缺陷 / Timeout forces defect
        fWinRatio := 0.0;               // 占比哨兵零（与真实占比可区分，看码）/ Sentinel ratio
        uCode := 16#0006_3034;          // 故障级：时长越限 / Fault: over duration
    ELSE
        _eVerdict := eDefect;           // 无样本保守缺陷 / Conservative defect without samples
        uCode := 16#0006_3033;          // 故障级：样本不足 / Fault: no samples
    END_IF
END_IF

(* 段 6｜出口装配 / Exit assembly *)
eVerdict := _eVerdict;                  // 判定输出 / Verdict output
IF NOT bRun THEN
    uCode := 16#0000_0000;              // 撤使能清码（可达解除）/ Run drop clears codes
END_IF
bError := (uCode >= 16#0006_3033) AND (uCode <= 16#0006_3035);  // 故障级码带判定 / Fault band check
uErrorId := uCode;                      // 码位单点写入 / Single write point
END_FUNCTION_BLOCK

(* ---- FB_DL_CalenderRollPress.st ---- *)
(*
  FB_DL_CalenderRollPress  —  辊压机辊隙/线压力顺控（双侧压下 + 厚度反馈） / Calender roll-gap and line-force sequencer with dual-side ram and thickness feedback
  分类 Category : DL_Process
  版本 Version  : 1.0.1
  来源 Source   : roadmap-li-p1 — 锂电极片辊压工站真缺口
  溯源 Origin   : 道莅 clean-room 实现；双侧压下同步 + 线压力建立 + 厚度窗监督为公开辊压工艺逻辑，未复制任何源码行
  功能 Function : 1) 四段顺控：eGapSet 双侧压下（左右辊隙均进目标容差带且同步偏差达标）→
                  eBarPress 线压力建立（fLinePressKn 进目标容差带）→ eRun 走带监视
                  （厚度窗 fThicknessUm 越窗即故障）→ eRelease 抬辊返回 → eDone；
                  2) 辊隙建立超时、线压力建立超时各自保护；3) 故障级单码 039F，
                  归因由 eCause 独立成员承载（R190）；4) 信息级 04C7 = 辊压循环完成沿；
                  5) 解除式全当拍量（R240）。
  接口 Interface: 输入双侧辊隙/线压力/厚度与两个时间量；输出状态/双侧镜像/厚度窗镜像/码。
                  抬辊计时 tonRun 复用 tGapTmo 常量（引脚预算取舍，非缺陷；若现场需独立抬辊超时，
                  下一版再增设 tReleaseTmo 引脚，引脚契约变更须走 MINOR 版本而非 PATCH）
  边界 Boundary : ① 组态闸：fGapTolMm <= 0.0、fLinePressTolKn <= 0.0、fGapSyncMaxMm <= 0.0、
                  fThicknessHiUm <= fThicknessLoUm、tGapTmo <= T#0S、tPressTmo <= T#0S
                  任一成立 → 039F 锁存；五个组态实数同时做 NaN 自反判（见 ②），
                  否则 NaN 参与 `<= 0.0` 判据时恒假 → 组态闸静默失效；
                  ② 浮点判据全部容差式（ABS 差 <= 容差），禁 = / <> 判等；
                  〔例外〕NaN 自反判 [x <> x] 与 Inf 差值自减判 [(x-x) <> (x-x)] 是浮点判等禁令的
                  唯一合法例外（R79），只许用于「非有限检测」，不得用于任何工程量比较；
                  机检 G6 已对自反式加白名单；
                  ③ 双侧同步偏差 |左-右| > fGapSyncMaxMm，仅在 eGapSet / eBarPress / eRun 且
                  bStart 为真时判定（相位窗 _bSyncWin）；eIdle / eRelease / eDone 辊缝机械张开，
                  偏差属正常工况不判 —— R281 返修：消除 eIdle 上电即报与 eRelease 收尾误锁；
                  ④ 三个 TON + 一个 R_TRIG 段 0 无条件每周期调用，IN 由相位派生；
                  ⑤ 故障相迁出唯一路径 = bReset 上升沿；
                  ⑥ 零全局耦合（无 GVL / 无 VAR_EXTERNAL / 无直接物理地址访问）。
  依赖 Depends  : Standard.library（TON / R_TRIG）
  码表 Error codes（Process 段 0005，故障窗口 039F / 信息窗口 04C7）:
    16#0005_039F 故障级：辊压故障总码（组态非法 / 辊隙超时 / 双侧失同步 / 线压力超时 / 厚度越窗），
                 锁存至 bReset 上升沿；归因见 eCause，不新增码位（派单硬约束单码）
    16#0005_04C7 信息级：辊压循环完成沿（抬辊完成进 eDone 单拍）
  修订历史 Revision :
    2026-11-19  v1.0.0  R43 首版（批次 1 · 序号 3）
    2026-11-19  v1.0.1  R45 返修（R281）：同步判据加相位窗 _bSyncWin，消除 eIdle/eRelease 误锁 039F；
                        组态闸补 NaN 自反判（组态 NaN 曾使闸静默失效）；头注释边界③改写、接口段补
                        tonRun 复用 tGapTmo 说明；引脚契约零变更（PATCH）
*)

TYPE E_DL_CrpState :
(
    eIdle     := 0,    // 未使能待启动 / Idle, waiting start
    eGapSet   := 10,   // 双侧压下建立辊隙 / Dual-side gap setting
    eBarPress := 20,   // 线压力建立 / Line force build-up
    eRun      := 30,   // 走带运行（厚度窗监督） / Running under thickness window
    eRelease  := 40,   // 抬辊返回 / Roll release
    eDone     := 50,   // 循环完成 / Done
    eFault    := 90    // 故障锁存相 / Fault latched phase
);
END_TYPE

TYPE E_DL_CrpCause :
(
    eNone       := 0,  // 无故障成因 / No cause
    eCfgIllegal := 1,  // 组态非法 / Illegal configuration
    eGapTmo     := 2,  // 辊隙建立超时 / Gap setting timeout
    eGapSync    := 3,  // 双侧失同步（偏差超限） / Dual-side out of sync
    ePressTmo   := 4,  // 线压力建立超时 / Line force timeout
    eThkDev     := 5   // 厚度越窗 / Thickness out of window
);
END_TYPE

FUNCTION_BLOCK FB_DL_CalenderRollPress
VAR_INPUT
    fGapLeftMm      : REAL := 0.0;      // 操作侧辊隙 [mm] / Operator-side roll gap
    fGapRightMm     : REAL := 0.0;      // 传动侧辊隙 [mm] / Drive-side roll gap
    fGapTargetMm    : REAL := 0.120;    // 目标辊隙 [mm]，域 > 0 / Target roll gap
    fGapTolMm       : REAL := 0.005;    // 辊隙容差带 [mm]，域 > 0 / Roll gap tolerance
    fGapSyncMaxMm   : REAL := 0.010;    // 双侧允许同步偏差 [mm]，域 > 0 / Dual-side sync limit
    fLinePressKn    : REAL := 0.0;      // 实测线压力 [kN/cm] / Measured line force
    fLinePressTgtKn : REAL := 12.0;     // 目标线压力 [kN/cm]，域 > 0 / Target line force
    fLinePressTolKn : REAL := 0.5;      // 线压力容差带 [kN/cm]，域 > 0 / Line force tolerance
    fThicknessUm    : REAL := 0.0;      // 实测极片厚度 [µm] / Measured electrode thickness
    fThicknessLoUm  : REAL := 100.0;    // 厚度窗下限 [µm] / Thickness low limit
    fThicknessHiUm  : REAL := 140.0;    // 厚度窗上限 [µm] / Thickness high limit
    tGapTmo         : TIME := T#10S;    // 辊隙建立超时 [ms]，域 > 0 / Gap timeout
    tPressTmo       : TIME := T#10S;    // 线压力建立超时 [ms]，域 > 0 / Force timeout
    bStart          : BOOL := FALSE;    // 启动命令（电平）[-] / Start command
    bReset          : BOOL := FALSE;    // 复位命令，上升沿清故障 [-] / Reset edge
END_VAR
VAR_OUTPUT
    eState          : E_DL_CrpState;    // 状态出口，段 6 单点映射 / State outlet
    eCause          : E_DL_CrpCause;    // 故障成因出口（R190） / Fault cause outlet
    fGapMeanMm      : REAL;             // 双侧辊隙均值 [mm] / Mean roll gap
    bGapOk          : BOOL;             // 辊隙达窗镜像 [-] / Gap in-window mirror
    bThkOk          : BOOL;             // 厚度在窗镜像 [-] / Thickness in-window mirror
    bCycleDone      : BOOL;             // 循环完成标志 [-] / Cycle done flag
    bError          : BOOL;             // 故障锁存标志 [-] / Fault latch flag
    nErrId          : UDINT;            // 事件码，0 = 无事件 / Event code
END_VAR
VAR
    _eState         : E_DL_CrpState := E_DL_CrpState.eIdle;   // 内部相位（CASE 唯一写入目标） / Internal phase
    _eCause         : E_DL_CrpCause := E_DL_CrpCause.eNone;   // 故障成因锁存（锁存量） / Latched cause
    tonGap          : TON;              // 辊隙建立计时，每周期无条件调用 / Gap timer
    tonPress        : TON;              // 线压力建立计时，每周期无条件调用 / Force timer
    tonRun          : TON;              // 抬辊计时，每周期无条件调用 / Release timer
    rtReset         : R_TRIG;           // 复位沿实例，每周期无条件调用 / Reset edge
    _fGapDev        : REAL;             // 双侧辊隙偏差 [mm]（当拍量） / Dual-side gap deviation
    _fGapErr        : REAL;             // 单侧辊隙对目标偏差 [mm]（当拍量） / Single-side gap error
    _bSyncWin       : BOOL;             // 双侧同步判据窗当拍量 [-]（单拍量，不入锁存清单） / Sync criterion window (per-scan)
    _bGapOk         : BOOL;             // 辊隙达窗当拍量 [-] / Gap verdict
    _bThkOk         : BOOL;             // 厚度在窗当拍量 [-] / Thickness verdict
    _bCfgBad        : BOOL;             // 组态非法当拍量 [-] / Config illegal
    _bFault         : BOOL;             // 故障锁存位（锁存量） / Latched fault bit
    _uFault         : UDINT;            // 故障码锁存（锁存量） / Latched fault code
    _uInfo          : UDINT;            // 信息码，每拍重算 / Transient info code
END_VAR

(* —— 段 0：沿实例与定时器无条件周期刷新 —— *)
_fGapDev := fGapLeftMm - fGapRightMm;                                          // 双侧辊隙偏差 / Dual-side deviation
_bSyncWin := bStart AND ((_eState = E_DL_CrpState.eGapSet)
                      OR (_eState = E_DL_CrpState.eBarPress)
                      OR (_eState = E_DL_CrpState.eRun));                      // 同步判据窗：仅在压下/建压/走带且启动电平在效时判同步 [-] / Sync window
_fGapErr := fGapLeftMm - fGapTargetMm;                                         // 操作侧对目标偏差 / Operator-side error
_bGapOk := (ABS(_fGapErr) <= fGapTolMm) AND (ABS(fGapRightMm - fGapTargetMm) <= fGapTolMm);   // 双侧均在容差带 / Both sides within tolerance
_bThkOk := (fThicknessUm >= fThicknessLoUm - 1.0E-6) AND (fThicknessUm <= fThicknessHiUm + 1.0E-6);  // 厚度容差窗 / Thickness window
_bCfgBad := (fGapTolMm <> fGapTolMm) OR (fLinePressTolKn <> fLinePressTolKn) OR (fGapSyncMaxMm <> fGapSyncMaxMm)
            OR (fThicknessLoUm <> fThicknessLoUm) OR (fThicknessHiUm <> fThicknessHiUm)   // NaN 自反判（禁令唯一例外 R79）/ NaN self-test
            OR (fGapTolMm <= 0.0) OR (fLinePressTolKn <= 0.0) OR (fGapSyncMaxMm <= 0.0)
            OR (fThicknessHiUm <= fThicknessLoUm) OR (tGapTmo <= T#0S) OR (tPressTmo <= T#0S);  // 组态非法当拍量 / Config illegal
rtReset(CLK := bReset);                                                        // 复位沿，每拍必调 / Reset edge
tonGap(IN := (_eState = E_DL_CrpState.eGapSet), PT := tGapTmo);                // 辊隙建立计时 / Gap timer
tonPress(IN := (_eState = E_DL_CrpState.eBarPress), PT := tPressTmo);          // 线压力建立计时 / Force timer
tonRun(IN := (_eState = E_DL_CrpState.eRelease), PT := tGapTmo);               // 抬辊计时（复用辊隙超时常量） / Release timer

(* —— 段 1：单拍量预清零（锁存量不入清单） —— *)
_uInfo := 16#0000_0000;            // 信息码每拍重算 / Info recomputed
fGapMeanMm := 0.0;                 // 辊隙均值缺省 0 / Mean gap default
bGapOk := FALSE;                   // 辊隙镜像缺省 FALSE / Gap flag default
bThkOk := FALSE;                   // 厚度镜像缺省 FALSE / Thickness flag default
bCycleDone := FALSE;               // 完成标志缺省 FALSE / Done default
nErrId := 16#0000_0000;            // 事件码缺省无事件 / Event code default

(* —— 段 2：复位沿（操作员复位语义：无条件清故障三件）+ 组态域闸 ——
   与段 4 分工：段 2 = 复位沿即刻清（不等解除式判据），段 4 = 解除式兜底判定；
   两段清同一三件，幂等无冲突（段 4 条件不成立时说明已被段 2 清毕，无需再动）。 *)
IF rtReset.Q THEN                              // rtReset.Q = 当拍量 / current scan
    _bFault := FALSE;                          // 清故障锁存位（锁存量） / Clear fault latch
    _uFault := 16#0000_0000;                   // 清故障锁存码（锁存量） / Clear fault code
    _eCause := E_DL_CrpCause.eNone;            // 清成因（锁存量） / Clear cause
    IF _eState = E_DL_CrpState.eFault THEN
        _eState := E_DL_CrpState.eIdle;        // 故障相迁出：回未使能 / Fault exit to idle
    END_IF
END_IF
IF _bCfgBad THEN                               // 组态域闸 / Config gate
    _uFault := 16#0005_039F;                   // 故障级：辊压故障总码 / Process fault code
    _bFault := TRUE;                           // 锁存置位 / Latch set
    bError := TRUE;                            // 故障标志同拍置位（R45 配对） / Error flag set same scan
    _eCause := E_DL_CrpCause.eCfgIllegal;      // 归因：组态非法 / Cause: illegal config
END_IF

(* —— 段 3：超时 / 失同步 / 厚度越窗（判据当拍量） —— *)
IF (NOT _bFault) AND tonGap.Q THEN             // 辊隙建立超时 / Gap timeout
    _uFault := 16#0005_039F;                   // 故障级：辊压故障总码 / Process fault code
    _bFault := TRUE;                           // 锁存置位 / Latch set
    bError := TRUE;                            // 故障标志同拍置位（R45 配对） / Error flag set same scan
    _eCause := E_DL_CrpCause.eGapTmo;          // 归因：辊隙超时 / Cause: gap timeout
END_IF
IF (NOT _bFault) AND _bSyncWin AND (ABS(_fGapDev) > fGapSyncMaxMm) THEN   // 仅同步窗内判（R281） / Only inside sync window
    _uFault := 16#0005_039F;                   // 故障级：辊压故障总码 / Process fault code
    _bFault := TRUE;                           // 锁存置位 / Latch set
    bError := TRUE;                            // 故障标志同拍置位（R45 配对） / Error flag set same scan
    _eCause := E_DL_CrpCause.eGapSync;         // 归因：失同步 / Cause: sync
END_IF
IF (NOT _bFault) AND tonPress.Q THEN           // 线压力建立超时 / Force timeout
    _uFault := 16#0005_039F;                   // 故障级：辊压故障总码 / Process fault code
    _bFault := TRUE;                           // 锁存置位 / Latch set
    bError := TRUE;                            // 故障标志同拍置位（R45 配对） / Error flag set same scan
    _eCause := E_DL_CrpCause.ePressTmo;        // 归因：线压力超时 / Cause: force timeout
END_IF
IF (NOT _bFault) AND (_eState = E_DL_CrpState.eRun) AND (NOT _bThkOk) THEN   // 走带期厚度越窗 / Thickness deviation
    _uFault := 16#0005_039F;                   // 故障级：辊压故障总码 / Process fault code
    _bFault := TRUE;                           // 锁存置位 / Latch set
    bError := TRUE;                            // 故障标志同拍置位（R45 配对） / Error flag set same scan
    _eCause := E_DL_CrpCause.eThkDev;          // 归因：厚度越窗 / Cause: thickness
END_IF

(* —— 段 4：故障解除式（R240；全当拍量）：rtReset.Q / NOT _bCfgBad / NOT tonGap.Q / NOT tonPress.Q ——
   解除式自证可满足（终审两式 1）：故障相内 _eState = eFault → tonGap.IN 与 tonPress.IN 恒假
   → 两 Q 恒假；操作员按复位时只需组态合法（NOT _bCfgBad），四因子即可同时为真 → 达式可满足、
   非 R152 恒假组合。刻意不追加 NOT _bSyncWin：故障相内 _bSyncWin 已恒假，追加即恒真冗余项；
   且复位后 _eState 回 eIdle → _bSyncWin 恒假 → 同步判据不复锁，解除可达性不依赖该因子。 *)
IF rtReset.Q AND (NOT _bCfgBad) AND (NOT tonGap.Q) AND (NOT tonPress.Q) THEN
    _bFault := FALSE;                          // 清故障锁存位（锁存量） / Clear fault latch
    _uFault := 16#0000_0000;                   // 清故障锁存码（锁存量） / Clear fault code
    _eCause := E_DL_CrpCause.eNone;            // 清成因（锁存量） / Clear cause
END_IF

(* —— 段 4A：故障锁存相位迁移闸 —— *)
IF _bFault AND (_eState <> E_DL_CrpState.eFault) THEN
    _eState := E_DL_CrpState.eFault;           // 锁存即入故障相 / Latch enters fault phase
END_IF

(* —— 段 5：相位机（CASE 全覆盖 + ELSE 兜底） —— *)
CASE _eState OF

E_DL_CrpState.eIdle:
    IF bStart AND (NOT _bFault) THEN           // 启动条件 / Start gate
        _eState := E_DL_CrpState.eGapSet;      // 进辊隙建立相 / Enter gap setting
    END_IF

E_DL_CrpState.eGapSet:
    IF _bGapOk THEN                            // 出口 1：双侧辊隙达窗 / Gap reached
        _eState := E_DL_CrpState.eBarPress;    // 进线压力相 / Enter force build-up
    ELSIF NOT bStart THEN                      // 出口 2：撤启动（R98 双出口） / Start released
        _eState := E_DL_CrpState.eRelease;     // 直接抬辊返回 / Go release
    END_IF

E_DL_CrpState.eBarPress:
    IF ABS(fLinePressKn - fLinePressTgtKn) <= fLinePressTolKn THEN   // 线压力达容差带 / Force reached band
        _eState := E_DL_CrpState.eRun;         // 进走带相 / Enter running
    ELSIF NOT bStart THEN                      // 撤启动：抬辊返回 / Start released
        _eState := E_DL_CrpState.eRelease;
    END_IF

E_DL_CrpState.eRun:
    IF NOT bStart THEN                         // 撤启动：进抬辊相 / Start released enters release
        _eState := E_DL_CrpState.eRelease;
    END_IF

E_DL_CrpState.eRelease:
    IF tonRun.Q THEN                           // 抬辊计时到 / Release elapsed
        _uInfo := 16#0005_04C7;                // 信息级：循环完成沿 / Info: cycle complete edge
        _eState := E_DL_CrpState.eDone;        // 进完成相 / Enter done
    END_IF

E_DL_CrpState.eDone:
    IF bStart THEN                             // 新循环上升请求 / New cycle request
        _eState := E_DL_CrpState.eGapSet;      // 直接进辊隙相 / Enter gap phase
    END_IF

E_DL_CrpState.eFault:
    ;                                          // 故障相：仅段 4 复位沿可迁出 / Only reset exits

ELSE
    _uFault := 16#0005_039F;                   // 故障级：非法相位兜底（归并总码） / Illegal phase fallback
    _bFault := TRUE;                           // 锁存置位 / Latch set
    bError := TRUE;                            // 故障标志同拍置位（R45 配对） / Error flag set same scan
    _eCause := E_DL_CrpCause.eCfgIllegal;      // 归因：相位非法归并组态 / Cause: phase illegal
    _eState := E_DL_CrpState.eFault;           // 强制回故障相 / Force fault phase

END_CASE

(* —— 段 6：出口单点映射（名实同源；锁存码回放） —— *)
fGapMeanMm := (fGapLeftMm + fGapRightMm) * 0.5;   // 双侧辊隙均值 / Mean roll gap
bGapOk := _bGapOk AND (NOT _bFault);              // 辊隙镜像 / Gap mirror
bThkOk := _bThkOk AND (NOT _bFault);              // 厚度镜像 / Thickness mirror
bCycleDone := (_eState = E_DL_CrpState.eDone);    // 完成标志 / Done flag
IF _bFault THEN
    nErrId := _uFault;                         // 故障锁存码回放 / Replay latched code
ELSE
    nErrId := _uInfo;                          // 信息码 / Transient info
END_IF
bError := _bFault;                             // 故障标志同源 / Flag from latch
eState := _eState;                             // 状态出口 / State outlet
eCause := _eCause;                             // 成因出口 / Cause outlet

END_FUNCTION_BLOCK

(* ---- FB_DL_CartonDenestPush.st ---- *)
(*
  FB_DL_CartonDenestPush  —  纸箱分离-推箱顺控 / Carton denesting and push sequence
  分类 Category : DL_Process
  码位 Code     : 16#06_0_B8
  段位说明      : R38 W7 预留 B6~BF 本轮正式启用，B7 格由 ElectrolyteFillCtrl 启用，本件启用 B8 格
  版本 Version  : 1.0.0
  来源 Source   : t2-7-packml — 成型上游分离供箱工艺待挖项
  溯源 Origin   : clean-room 实现，未复制任何源码行
                  （与 FB_DL_CartonErectSeq / CartonErectorStation 分工：那族管开箱成型，本件是成型上游的分离供箱）
  功能 Function : 1) 七相顺控 Idle→LevelChk→VacPick→SepLift→Push→PushRet→Drop→Done：
                  料位联锁 → 真空吸取顶箱 → 分离缸提升 → 推杆推箱 → 推杆缩回 → 落箱放行；
                  2) 双联锁内置：推箱须「真空保持 AND 箱在位」双确认，联锁不满足只等待不故障；
                  3) 双料位联锁：低料位且无高料位判料仓耗尽（信息级等待，不启动新周期）；
                  4) 段超时升级：五段各配独立超时 TON，超时锁故障（安全侧全停）。
  边界 Boundary : ① 真空接口契约：iEjector.fPressure 为负压值，吸取确认深度 = −fPressure；
                  ② 组态域闸覆盖全部参与换算引脚（R151）；
                  ③ R228-A 达标声明：五只超时 TON 均单相独占（IN 为单相等式），跨相迁移拍 IN 必断；
                  ④ R228-B 达标声明：eFault 迁出 = rtReset.Q（输入引脚，恒可达），逐字写于此；
                  ⑤ 气缸命令经 I_DL_Cylinder 方法单发下发（方法内受理去重，重复调用无害）；
                  ⑥ CASE 全态覆盖 + ELSE 兜底置 Fault。
  依赖 Depends  : I_DL_Cylinder（×2 注入：分离缸/推箱缸，不实例化）；
                  I_DL_VacuumGenerator（注入，不实例化；FB_DL_VacuumEjector 为典型实现）；
                  段序语义对齐 FB_DL_StepSequencer（已注册，不实例化）
  码表 Error codes（本件格 06_0_B8，子码步进 +0x100）:
    16#0006_01B8 信息级：供箱周期完成（Done 相）
    16#0006_02B8 故障级：组态非法（吸取深度/常压阈/超时域非法），锁存至复位
    16#0006_03B8 故障级：段超时升级（五段独立计时），锁存至复位
    16#0006_04B8 故障级：注入件故障（分离缸/推箱缸/真空 bFault），锁存至复位
    16#0006_05B8 信息级：料仓耗尽（低料位且无高料位，等待补料，不置故障）
    16#0006_06B8 信息级：推箱双联锁等待（真空/箱在位未齐，不置故障）
    16#0006_07B8 故障级：状态机落 ELSE 兜底（非法相位 ID）

  修订历史 Revision :
    2026-11-19  v1.0.0  R39 首版（批次 4 · 序号 16）
*)

TYPE E_DL_DenestState :
(
    eIdle     := 0,    // 空闲：等启动指令 / Idle, waiting for start
    eLevelChk := 10,   // 料位检查：联锁判定 / Level check interlock
    eVacPick  := 20,   // 真空吸取：建立吸取真空 / Vacuum pick, establish holding vacuum
    eSepLift  := 30,   // 分离提升：分离缸伸出 / Separate lift, separator cylinder extend
    ePush     := 40,   // 推箱：推杆伸出（双联锁内） / Push, pusher extend under dual interlock
    ePushRet  := 50,   // 推杆缩回 / Pusher retract
    eDrop     := 60,   // 落箱：分离缸缩回 + 破真空 / Drop, separator retract and blow-off
    eDone     := 70,   // 完成：周期落定 / Done
    eFault    := 90    // 故障：组态/超时/注入件锁定 / Fault, latched
);
END_TYPE

FUNCTION_BLOCK FB_DL_CartonDenestPush
VAR_INPUT
    bStart       : BOOL := FALSE;      // 启动指令（上升沿）/ Start command
    bBoxAtPick   : BOOL := FALSE;      // 取箱位有箱反馈 [-] / Box present at pick position
    bBoxMagHigh  : BOOL := FALSE;      // 料仓高料位反馈 [-] / Magazine high-level feedback
    bBoxMagLow   : BOOL := FALSE;      // 料仓低料位反馈 [-] / Magazine low-level feedback
    fVacPickKpa  : REAL := 40.0;       // 吸取确认深度 [kPa]，域 > 0 / Pick confirmation vacuum depth
    fAtmVacKpa   : REAL := 5.0;        // 落箱常压确认阈 [kPa]，域 >= 0 / Drop atmospheric threshold
    tStepTimeout : TIME := T#5S;       // 单段超时 [ms]，域 > 0 / Per-step timeout
    bReset       : BOOL := FALSE;      // 复位（eFault 迁出唯一沿）/ Reset, sole fault exit edge
END_VAR
VAR_OUTPUT
    bCycleDone   : BOOL;               // 供箱周期完成 / Cycle done
    nStep        : INT;                // 当前步号 [0..4]（0=吸取 1=提升 2=推箱 3=缩回 4=落箱）/ Step index
    bPushPermit  : BOOL;               // 推箱双联锁满足 [-] / Push dual interlock satisfied
    bMagEmpty    : BOOL;               // 料仓耗尽指示 [-] / Magazine empty indicator
    nErrId       : UDINT;              // 事件码，0 = 无事件 / Event code
    eState       : E_DL_DenestState;   // 状态出口，段尾单点映射 / State outlet
END_VAR
VAR_IN_OUT
    iSepCyl   : I_DL_Cylinder;         // 分离缸引用（注入，不实例化）/ Separator cylinder reference
    iPushCyl  : I_DL_Cylinder;         // 推箱缸引用（注入，不实例化）/ Pusher cylinder reference
    iEjector  : I_DL_VacuumGenerator;  // 真空发生器引用（注入，不实例化）/ Vacuum generator reference
END_VAR
VAR
    tonVacTo  : TON;                   // 吸取段超时（单相独占）/ Pick timeout, single phase
    tonSepTo  : TON;                   // 提升段超时（单相独占）/ Lift timeout, single phase
    tonPushTo : TON;                   // 推箱段超时（单相独占）/ Push timeout, single phase
    tonRetTo  : TON;                   // 缩回段超时（单相独占）/ Retract timeout, single phase
    tonDropTo : TON;                   // 落箱段超时（单相独占）/ Drop timeout, single phase
    tonWch    : TON;                   // 故障观察窗，自复位 / Fault watch window, self-resetting
    rtStart   : R_TRIG;                // 启动上升沿 / Start rising edge
    rtReset   : R_TRIG;                // 复位上升沿 / Reset rising edge
    _eState   : E_DL_DenestState := E_DL_DenestState.eIdle;   // 内部相位（CASE 唯一写入目标）/ Internal phase
    _rVacDep  : REAL;                  // 真空深度暂存 [kPa] / Vacuum depth scratch
    _bVacOk   : BOOL;                  // 吸取确认标志 / Pick confirmed flag
    _bVacRel  : BOOL;                  // 常压确认标志 / Atmospheric confirmed flag
    _uFault   : UDINT;                 // 故障码锁存 / Latched fault code
    _uInfo    : UDINT;                 // 信息码，每拍重算 / Info code
    _bFault   : BOOL;                  // 故障锁存位 / Latched fault bit
    _bCfgBad  : BOOL;                  // 组态非法聚合 / Configuration invalid aggregate
END_VAR
VAR CONSTANT
    DL_CDP_WATCH_PT : TIME := T#2S;   // 故障观察窗 [ms]，自复位 / Fault watch window
    DL_CDP_INF_CAP  : REAL := 1.0E15; // 非有限值筛查幅值上限 / Non-finite screening cap
END_VAR

(* —— 段 0：定时器与边沿无条件周期刷新（R182：调用语句不得置于 IF/CASE 内） —— *)
rtStart(CLK := bStart);                                                // 启动沿刷新，每拍必调
rtReset(CLK := bReset);                                                // 复位沿刷新，每拍必调
tonWch(IN := (NOT tonWch.Q), PT := DL_CDP_WATCH_PT);                   // 观察窗自复位（表达式入参）
tonVacTo(IN := (_eState = E_DL_DenestState.eVacPick), PT := tStepTimeout);   // 吸取超时（单相独占）
tonSepTo(IN := (_eState = E_DL_DenestState.eSepLift), PT := tStepTimeout);   // 提升超时（单相独占）
tonPushTo(IN := (_eState = E_DL_DenestState.ePush), PT := tStepTimeout);     // 推箱超时（单相独占）
tonRetTo(IN := (_eState = E_DL_DenestState.ePushRet), PT := tStepTimeout);   // 缩回超时（单相独占）
tonDropTo(IN := (_eState = E_DL_DenestState.eDrop), PT := tStepTimeout);     // 落箱超时（单相独占）

(* —— 段 1：单拍量预清零（锁存量 _uFault/_bFault 不入清单，R187①） —— *)
_uInfo := 16#0000_0000;             // 信息码每拍重算
bCycleDone := FALSE;                // 完成出口缺省 FALSE（Done 相单点置位）
bPushPermit := FALSE;               // 双联锁出口缺省 FALSE（段 5 单点重写）
_bCfgBad := FALSE;                  // 组态非法预清零
nErrId := 16#0000_0000;             // 事件码缺省无事件

(* —— 段 2：组态域闸（覆盖全部参与判据换算的引脚，R151） —— *)
IF (fVacPickKpa <> fVacPickKpa) OR (fVacPickKpa <= 0.0) OR (ABS(fVacPickKpa) > DL_CDP_INF_CAP)
   OR (fAtmVacKpa < 0.0) OR (TIME_TO_DINT(tStepTimeout) <= 0) THEN
    _bCfgBad := TRUE;               // 吸取深度/常压阈/超时非法
END_IF

(* —— 段 3：eFault 迁出沿（R228-B：rtReset.Q 为输入引脚，恒可达） —— *)
IF rtReset.Q THEN
    _bFault := FALSE;               // 清故障锁存位
    _uFault := 16#0000_0000;
    IF _eState = E_DL_DenestState.eFault THEN
        _eState := E_DL_DenestState.eIdle;      // 故障相迁出：回空闲
    END_IF
END_IF

(* —— 段 4：过程量只读采集与判据 —— *)
_rVacDep := -iEjector.fPressure;                // 真空深度 = 负压反馈取反 [kPa]（接口契约：负值=真空）
_bVacOk := _rVacDep >= fVacPickKpa;             // 吸取确认（每拍重算）
_bVacRel := _rVacDep <= fAtmVacKpa;             // 常压确认（每拍重算）
bMagEmpty := bBoxMagLow AND (NOT bBoxMagHigh);  // 料仓耗尽派生（每拍重算）

(* —— 段 5：相位机（只做迁移与单发命令；出口在段 7） —— *)
CASE _eState OF

E_DL_DenestState.eIdle:
    IF rtStart.Q AND _bCfgBad THEN
        _uFault := 16#0006_02B8;            // 故障级：组态非法
        _bFault := TRUE;
        _eState := E_DL_DenestState.eFault;
    ELSIF rtStart.Q AND bMagEmpty THEN
        _uInfo := 16#0006_05B8;             // 信息级：料仓耗尽等待补料（不启动周期）
    ELSIF rtStart.Q AND (NOT _bCfgBad) THEN
        _eState := E_DL_DenestState.eLevelChk;  // 进料位检查相
    END_IF

E_DL_DenestState.eLevelChk:
    IF (iSepCyl.bFault OR iPushCyl.bFault OR iEjector.bFault) THEN
        _uFault := 16#0006_04B8;            // 故障级：注入件故障
        _bFault := TRUE;
        iEjector.CmdStop();                 // 安全侧全停
        _eState := E_DL_DenestState.eFault;
    ELSIF bMagEmpty THEN
        _uInfo := 16#0006_05B8;             // 信息级：料仓耗尽（退回空闲等补料）
        _eState := E_DL_DenestState.eIdle;
    ELSE
        iEjector.CmdEvacuate();             // 单发吸取指令
        _eState := E_DL_DenestState.eVacPick;   // 进吸取相
    END_IF

E_DL_DenestState.eVacPick:
    IF (iSepCyl.bFault OR iPushCyl.bFault OR iEjector.bFault) THEN
        _uFault := 16#0006_04B8;
        _bFault := TRUE;
        iEjector.CmdStop();
        _eState := E_DL_DenestState.eFault;
    ELSIF tonVacTo.Q THEN
        _uFault := 16#0006_03B8;            // 故障级：吸取段超时
        _bFault := TRUE;
        iEjector.CmdStop();
        _eState := E_DL_DenestState.eFault;
    ELSIF _bVacOk AND tonWch.Q THEN
        iSepCyl.CmdExtend();                // 单发提升指令
        _eState := E_DL_DenestState.eSepLift;   // 进提升相
    END_IF

E_DL_DenestState.eSepLift:
    IF (iSepCyl.bFault OR iPushCyl.bFault OR iEjector.bFault) THEN
        _uFault := 16#0006_04B8;
        _bFault := TRUE;
        iSepCyl.CmdStop();
        iEjector.CmdStop();
        _eState := E_DL_DenestState.eFault;
    ELSIF tonSepTo.Q THEN
        _uFault := 16#0006_03B8;            // 故障级：提升段超时
        _bFault := TRUE;
        iSepCyl.CmdStop();
        _eState := E_DL_DenestState.eFault;
    ELSIF iSepCyl.bExtended THEN
        _eState := E_DL_DenestState.ePush;  // 提升到位：进推箱相
    END_IF

E_DL_DenestState.ePush:
    bPushPermit := _bVacOk AND bBoxAtPick;  // 双联锁派生出口（每拍重算）
    IF (iSepCyl.bFault OR iPushCyl.bFault OR iEjector.bFault) THEN
        _uFault := 16#0006_04B8;
        _bFault := TRUE;
        iPushCyl.CmdStop();
        _eState := E_DL_DenestState.eFault;
    ELSIF tonPushTo.Q THEN
        _uFault := 16#0006_03B8;            // 故障级：推箱段超时
        _bFault := TRUE;
        iPushCyl.CmdStop();
        _eState := E_DL_DenestState.eFault;
    ELSIF NOT bPushPermit THEN
        _uInfo := 16#0006_06B8;             // 信息级：双联锁等待（不置故障）
    ELSE
        iPushCyl.CmdExtend();               // 联锁满足：单发推箱
        IF iPushCyl.bExtended THEN
            iPushCyl.CmdRetract();          // 推到位即单发缩回
            _eState := E_DL_DenestState.ePushRet;   // 进缩回相
        END_IF
    END_IF

E_DL_DenestState.ePushRet:
    IF (iSepCyl.bFault OR iPushCyl.bFault OR iEjector.bFault) THEN
        _uFault := 16#0006_04B8;
        _bFault := TRUE;
        iPushCyl.CmdStop();
        _eState := E_DL_DenestState.eFault;
    ELSIF tonRetTo.Q THEN
        _uFault := 16#0006_03B8;            // 故障级：缩回段超时
        _bFault := TRUE;
        iPushCyl.CmdStop();
        _eState := E_DL_DenestState.eFault;
    ELSIF iPushCyl.bRetracted THEN
        iSepCyl.CmdRetract();               // 单发分离缸缩回
        iEjector.CmdBlowOff();              // 单发破真空落箱
        _eState := E_DL_DenestState.eDrop;  // 进落箱相
    END_IF

E_DL_DenestState.eDrop:
    IF (iSepCyl.bFault OR iPushCyl.bFault OR iEjector.bFault) THEN
        _uFault := 16#0006_04B8;
        _bFault := TRUE;
        iSepCyl.CmdStop();
        _eState := E_DL_DenestState.eFault;
    ELSIF tonDropTo.Q THEN
        _uFault := 16#0006_03B8;            // 故障级：落箱段超时
        _bFault := TRUE;
        _eState := E_DL_DenestState.eFault;
    ELSIF iSepCyl.bRetracted AND _bVacRel THEN
        _eState := E_DL_DenestState.eDone;  // 缩回 + 常压双确认：进完成相
    END_IF

E_DL_DenestState.eDone:
    bCycleDone := TRUE;                     // 完成出口（Done 相每拍重申）
    _uInfo := 16#0006_01B8;                 // 信息级：周期完成
    IF NOT bStart THEN
        _eState := E_DL_DenestState.eIdle;  // 指令撤销：回空闲
    END_IF

E_DL_DenestState.eFault:
    ;                                       // 故障相：等复位沿（段 3 承载迁出）

ELSE
    _uFault := 16#0006_07B8;                // 故障级：非法相位 ID 兜底
    _bFault := TRUE;
    _eState := E_DL_DenestState.eFault;     // 强制回故障相

END_CASE

(* —— 段 6：出口单点映射（名实同源；锁存码回放，禁同拍抹除） —— *)
IF _eState = E_DL_DenestState.eVacPick THEN
    nStep := 0;                             // 步号 0：吸取
ELSIF _eState = E_DL_DenestState.eSepLift THEN
    nStep := 1;                             // 步号 1：提升
ELSIF _eState = E_DL_DenestState.ePush THEN
    nStep := 2;                             // 步号 2：推箱
ELSIF _eState = E_DL_DenestState.ePushRet THEN
    nStep := 3;                             // 步号 3：缩回
ELSIF _eState = E_DL_DenestState.eDrop THEN
    nStep := 4;                             // 步号 4：落箱
ELSE
    nStep := -1;                            // Idle/LevelChk/Done/Fault：无有效步号
END_IF
IF _bFault THEN
    nErrId := _uFault;                      // 故障锁存码回放（不在故障相按当下输入重推）
    bCycleDone := FALSE;                    // 故障相完成出口强制 FALSE（安全侧）
    bPushPermit := FALSE;                   // 故障相联锁出口强制 FALSE（安全侧）
ELSE
    nErrId := _uInfo;                       // 信息码
END_IF
eState := _eState;                          // 状态出口单点映射

END_FUNCTION_BLOCK

(* ---- FB_DL_CartonErectorStation.st ---- *)
//==============================================================================
// 功能块：FB_DL_CartonErectorStation ｜ 中文名称：开箱（Carton Erector）工站模板
// 所属子库：DL_Process ｜ 版本：v1.0.1 ｜ 兼容：CODESYS V3.5+ / TwinCAT 3 / 汇川 InoProShop
// 功能描述：开箱工站七态九步骨架——七态 = 就绪/送箱坯/开箱/折底/插底/
//           封压/推出（外加 eIdle/eFault 两态不入工作态计数），九步 =
//           步进引擎步号 0..8（吸箱坯下降/吸持/提升/撑箱开箱/折前底翼/
//           折后底翼/插底翼锁底/压底整形/推出），步完成由本件按反馈与
//           驻留判据装配，步超时由 FB_DL_StepSequencer 统一监控（DL_Base
//           组合调用，接口引脚契约与 FB_DL_ElectrolyteDosingSeq 同口径）。
//           步号-相位映射表：0/1/2 → eFeeding（送坯三步）、3 → eOpening、
//           4/5/6 → eFolding、7 → eSealing、8 → eEjecting、bDone → eDone。
// 开源溯源 (Origin)：道莅原创实现（参考 ISA-88 相-步骤语义与开箱成型机工程惯例 分类与参数域）
// 单位表：计数[次] / 时间[ms] / 阀输出[—]
// 错误码表：16#0005_01F4 信息级（成型完成放行：eDone 相进入，不置
//           bError）/ 16#0005_01F5 信息级（开箱到位提示：撑箱步完成，
//           关键节点可观测，不置 bError）/ 16#0005_0333 故障级（组态
//           非法：步超时表为 0 或箱坯 absent 且强行启动，置 bError）/
//           16#0005_0334 故障级（步超时：步进引擎判超时，锁存，置
//           bError——该场景不可由 0333 的组态类判据观测，属执行机构
//           独立域）/ 16#0005_0335 故障级兜底（状态机落 ELSE 或非法
//           状态，置 bError 并全输出断）
// 状态机：E_DL_CartonPhase（九态：eIdle=0 / eReady=10 / eFeeding=20 /
//           eOpening=30 / eFolding=40 / eSealing=50 / eEjecting=60 /
//           eDone=70 / eFault=99；工作态七态 = eReady..eDone），CASE
//           含 ELSE 兜底，ELSE 置 0335 并全输出断
// 边界行为：① 组态非法（任一步超时为 0）→ 故障态锁存，bReset 复位；
//           ② bAbort → 两段化照 §4 修复件样板：真空/输出立即断，推出
//           缸保持不动，等运行条件消失回空闲；③ 步完成判据：反馈优先
//           （bXxxFb），无反馈步用驻留时间兜底；④ eDone 等启动撤销回
//           空闲（同拍重启防抖，R39 范式）；⑤ 未启动/故障全输出断
//           （真空、缸、推出全撤）；⑥ 安全侧 = abort 拍不得出现关阀
//           输出置位以外的任何缸动作（机检断言：abort 拍仅真空断）。
// 依赖纪律：Process → Level 0 组合调用合法——步进引擎组合调用
//           FB_DL_StepSequencer（DL_Base，接口已核实），全库单调用点
//           （每拍恰好调用一次，防双调用边沿竞态）。
// 修订历史：v1.0.0 2026-11-17 首版（R24 派单 · ROADMAP P0 §652）
//           v1.0.1 2026-11-17 R24 终审修复（R106 第一档，契约不变）：原
//           fbSeq.bReset 恒 FALSE，而步进引擎 bError 为锁存型
//          （eState = eFault，仅 bReset 上升沿清除），步超时后工站故障
//           恢复条件 NOT fbSeq.bError 永不满足 → 故障恢复死锁；修复为
//           仅在工站 eFault 相透传 bReset，非故障相禁透传（防运行中误清
//           步进器致相位-步号失配）。引脚契约、码位、枚举不变。
//==============================================================================

(*------------------------------------------------------------------------------
 * 枚举: E_DL_CartonPhase（归属本功能块，同文件发布，全库唯一定义）
 * 含义: 开箱工站相位，与步进器步号映射（0/1/2→eFeeding、3→eOpening、
 *       4/5/6→eFolding、7→eSealing、8→eEjecting）。
 *-----------------------------------------------------------------------------*)
TYPE E_DL_CartonPhase :
(
    eIdle     := 0,   // 空闲：等启动 / Idle, awaiting start
    eReady    := 10,  // 就绪：箱坯在位确认窗（步 0 吸箱坯下降） / Ready, blank presence window, step 0
    eFeeding  := 20,  // 送箱坯：吸持提升（步 1/2） / Feeding, vacuum and lift, steps 1 and 2
    eOpening  := 30,  // 开箱：撑箱开箱（步 3） / Opening, case spreader, step 3
    eFolding  := 40,  // 折底：折前后底翼与插底锁底（步 4/5/6） / Folding, bottom flaps and tuck, steps 4 to 6
    eSealing  := 50,  // 封压：压底整形（步 7） / Sealing, bottom press, step 7
    eEjecting := 60,  // 推出：成品推出（步 8） / Ejecting, product push-out, step 8
    eDone     := 70,  // 完成：放行，等启动撤销 / Done, released, awaiting start drop
    eFault    := 99   // 故障：组态/步超时/非法状态 / Fault, config, step timeout or illegal state
);
END_TYPE

FUNCTION_BLOCK FB_DL_CartonErectorStation
VAR_INPUT
    bStart       : BOOL;                    // 启动请求 [—]，上升沿生效 / Start request, rising edge
    bAbort       : BOOL;                    // 中止请求 [—]，任意拍生效 / Abort request, effective on any scan
    bReset       : BOOL;                    // 故障复位 [—]，上升沿清锁存 / Fault reset, rising edge clears latches
    bBlankPresent: BOOL;                    // 箱坯在位 [—] / Carton blank present
    bVacuumFb    : BOOL;                    // 吸持真空反馈 [—] / Vacuum feedback
    bLiftFb      : BOOL;                    // 提升到位反馈 [—] / Lift-in-position feedback
    bOpenFb      : BOOL;                    // 开箱到位反馈 [—] / Spreader-in-position feedback
    bFoldFb      : BOOL;                    // 折翼到位反馈 [—] / Flap-in-position feedback
    bTuckFb      : BOOL;                    // 插底到位反馈 [—] / Tuck-in-position feedback
    bPressFb     : BOOL;                    // 压底到位反馈 [—] / Press-in-position feedback
    bEjectFb     : BOOL;                    // 推出到位反馈 [—] / Eject-in-position feedback
    tDwell       : TIME  := T#200MS;        // 无反馈步驻留兜底 [ms]，须 > 0 / Dwell fallback for feedback-less steps [ms]
END_VAR
VAR_OUTPUT
    ePhase       : E_DL_CartonPhase;        // 工站相位 [—] / Station phase
    bVacuumOn    : BOOL;                    // 吸持真空输出 [—] / Vacuum output
    bFeedOut     : BOOL;                    // 送箱坯下降输出 [—] / Blank-feed output
    bOpenOut     : BOOL;                    // 开箱缸输出 [—] / Spreader output
    bFoldOut     : BOOL;                    // 折翼缸输出 [—] / Flap cylinder output
    bTuckOut     : BOOL;                    // 插底缸输出 [—] / Tuck cylinder output
    bPressOut    : BOOL;                    // 压底缸输出 [—] / Press cylinder output
    bEjectOut    : BOOL;                    // 推出缸输出 [—] / Eject cylinder output
    eErr         : UDINT;                   // 错误码，0 = 无错，码位 16#0005_01F4 起信息级、16#0005_0333 起故障级（分带见错误码表） / Error code, 0 = no error, band info/fault per the code table
    bError       : BOOL;                    // 故障级标志，仅故障级错误置位 / Fault-class flag, set only on fault-level codes
    bValid       : BOOL;                    // 输出可用标志 / Outputs usable flag
END_VAR
VAR
    fbSeq        : FB_DL_StepSequencer;     // 步进引擎（Level 0 组合调用，单调用点） / Step engine, Level 0 composition, single call site
    fbDwellT     : TON;                     // 无反馈步驻留兜底计时（每拍无条件刷新）[ms] / Dwell fallback timer, refreshed unconditionally
    fbStart      : R_TRIG;                  // 启动沿检测（待机/故障分支同样无条件刷新） / Start edge detector, refreshed unconditionally
    _ePhase      : E_DL_CartonPhase := E_DL_CartonPhase.eIdle; // 当前相位 / Current phase
    _abStepDone  : ARRAY[0..15] OF BOOL;    // 步完成信号（本件按判据维护） / Step-done levels, maintained by this FB
    _auStepTimeout: ARRAY[0..15] OF TIME;   // 每步超时 [ms]，0 = 不监控 / Per-step timeout [ms], zero = not monitored
    _bSeqStart   : BOOL;                    // 步进器启动沿请求（单调用点输入） / Sequencer start edge request
    _bCfgBad     : BOOL;                    // 组态非法锁存 / Illegal config latch
    _bAbortStage : UINT;                    // 中止段号 [—]，0 = 无 / 1 = 输出已断 / Abort stage, zero none, one outputs cut
    _bInfoOpen   : BOOL;                    // 开箱到位信息当拍标志 / Opening info flag of this scan
    _bInfoDone   : BOOL;                    // 完成信息当拍标志 / Done info flag of this scan
    _bIllegal    : BOOL;                    // 非法状态标志 / Illegal state flag
    _bInit       : BOOL := FALSE;           // 首扫标志，初值 FALSE 取非判定 / First-scan flag, tested negated
END_VAR
VAR CONSTANT
    DL_CES_TO_FEED : TIME := T#3S;          // 步 0 吸箱坯超时 [ms] / Step 0 timeout [ms]
    DL_CES_TO_VAC  : TIME := T#2S;          // 步 1 吸持超时 [ms] / Step 1 timeout [ms]
    DL_CES_TO_LIFT : TIME := T#3S;          // 步 2 提升超时 [ms] / Step 2 timeout [ms]
    DL_CES_TO_OPEN : TIME := T#4S;          // 步 3 开箱超时 [ms] / Step 3 timeout [ms]
    DL_CES_TO_FOLD : TIME := T#3S;          // 步 4 折前底翼超时 [ms] / Step 4 timeout [ms]
    DL_CES_TO_FOLD2: TIME := T#3S;          // 步 5 折后底翼超时 [ms] / Step 5 timeout [ms]
    DL_CES_TO_TUCK : TIME := T#3S;          // 步 6 插底超时 [ms] / Step 6 timeout [ms]
    DL_CES_TO_PRESS: TIME := T#2S;          // 步 7 压底超时 [ms] / Step 7 timeout [ms]
    DL_CES_TO_EJCT : TIME := T#4S;          // 步 8 推出超时 [ms] / Step 8 timeout [ms]
END_VAR

(*------------------------------------------------------------------------------
 * 段 1｜每拍预置：全输出先断（安全侧），单拍标志预清零
 *      All outputs cleared first, fail-safe, one-shot flags pre-cleared
 *-----------------------------------------------------------------------------*)
bVacuumOn := FALSE;                      // 真空输出先清（安全侧） / Vacuum cleared first
bFeedOut  := FALSE;                      // 送坯输出先清 / Feed output cleared first
bOpenOut  := FALSE;                      // 开箱输出先清 / Spreader cleared first
bFoldOut  := FALSE;                      // 折翼输出先清 / Flap cleared first
bTuckOut  := FALSE;                      // 插底输出先清 / Tuck cleared first
bPressOut := FALSE;                      // 压底输出先清 / Press cleared first
bEjectOut := FALSE;                      // 推出输出先清 / Eject cleared first
eErr   := 16#0000_0000;                  // 错误码每拍重算 / Error code recomputed
bError := FALSE;                         // 故障标志每拍重算 / Fault flag recomputed
bValid := FALSE;                         // 可用标志每拍重算 / Usable flag recomputed
_bInfoOpen := FALSE;                     // 开箱信息预清零 / Opening info pre-cleared
_bInfoDone := FALSE;                     // 完成信息预清零 / Done info pre-cleared
_bIllegal  := FALSE;                     // 非法状态预清零 / Illegal flag pre-cleared
_bSeqStart := FALSE;                     // 步进器启动沿请求预清零 / Sequencer start request pre-cleared

(*------------------------------------------------------------------------------
 * 段 2｜首扫初始化：步超时表一次装配
 *      First-scan initialisation, the timeout table assembled once
 *-----------------------------------------------------------------------------*)
IF NOT _bInit THEN
    _ePhase := E_DL_CartonPhase.eIdle;   // 相位空闲起步 / Phase starts idle
    _auStepTimeout[0] := DL_CES_TO_FEED; // 步 0 超时 / Step 0 timeout
    _auStepTimeout[1] := DL_CES_TO_VAC;  // 步 1 超时 / Step 1 timeout
    _auStepTimeout[2] := DL_CES_TO_LIFT; // 步 2 超时 / Step 2 timeout
    _auStepTimeout[3] := DL_CES_TO_OPEN; // 步 3 超时 / Step 3 timeout
    _auStepTimeout[4] := DL_CES_TO_FOLD; // 步 4 超时 / Step 4 timeout
    _auStepTimeout[5] := DL_CES_TO_FOLD2; // 步 5 超时 / Step 5 timeout
    _auStepTimeout[6] := DL_CES_TO_TUCK; // 步 6 超时 / Step 6 timeout
    _auStepTimeout[7] := DL_CES_TO_PRESS; // 步 7 超时 / Step 7 timeout
    _auStepTimeout[8] := DL_CES_TO_EJCT; // 步 8 超时 / Step 8 timeout
    _auStepTimeout[9] := T#0MS;          // 步 9 及以后不监控 / Steps 9 and beyond not monitored
    _bCfgBad := FALSE;                   // 组态锁存清零 / Config latch cleared
    _bAbortStage := 0;                   // 中止段号从零起步 / Abort stage starts at zero
    _bInit := TRUE;                      // 首扫只做一次 / The first scan runs once
END_IF

(*------------------------------------------------------------------------------
 * 段 3｜组态闸 + 沿检测 + 驻留计时无条件刷新（R40：CASE 之外每拍必调）
 *      Config gate plus unconditional refresh per R40
 *-----------------------------------------------------------------------------*)
fbStart(CLK := bStart);                  // 启动沿检测 / Start edge detection
fbDwellT(IN := (_ePhase = E_DL_CartonPhase.eReady), PT := tDwell); // 步 0 吸箱坯下降驻留窗（进相即起算） / Step 0 feed-down dwell window, restarts on phase entry
IF (tDwell <= T#0MS) OR (_auStepTimeout[0] <= T#0MS)
   OR (_auStepTimeout[3] <= T#0MS) OR (_auStepTimeout[8] <= T#0MS) THEN
    _bCfgBad := TRUE;                    // 步超时表/驻留窗非法锁存（关键步抽查） / Timeout table and dwell domains latched, key steps sampled
END_IF

(*------------------------------------------------------------------------------
 * 段 4｜中止入口（输出立即断，机构位置保持）与复位
 *      Abort entry, outputs cut immediately, mechanisms held
 *-----------------------------------------------------------------------------*)
IF bAbort AND (_bAbortStage = 0)
   AND (_ePhase <> E_DL_CartonPhase.eIdle) AND (_ePhase <> E_DL_CartonPhase.eFault) THEN
    _bAbortStage := 1;                   // 进中止段（输出断、位置保持） / Enter abort stage, outputs cut, positions held
END_IF
IF _bAbortStage = 1 THEN
    IF (NOT bStart) THEN
        _bAbortStage := 0;               // 启动撤销回空闲 / Start dropped, back to idle
        _ePhase := E_DL_CartonPhase.eIdle; // 相位回空闲 / Phase back to idle
    END_IF
END_IF
IF bReset THEN
    _bCfgBad := FALSE;                   // 复位清组态锁存 / Reset clears the config latch
END_IF

(*------------------------------------------------------------------------------
 * 段 5｜步进器单调用点与步完成判据装配（每拍恰好一次）
 *      Single sequencer call site and step-done assembly
 *-----------------------------------------------------------------------------*)
_bSeqStart := fbStart.Q AND (_ePhase = E_DL_CartonPhase.eIdle)
              AND (NOT _bCfgBad) AND bBlankPresent; // 启动沿（空闲且组态合法且箱坯在位） / Start edge in idle with legal config and blank present
IF (_ePhase <> E_DL_CartonPhase.eIdle) AND (_ePhase <> E_DL_CartonPhase.eFault)
   AND (_bAbortStage = 0) THEN
    _abStepDone[0] := fbDwellT.Q;        // 步 0 完成：吸箱坯下降驻留窗满 / Step 0 done, feed-down dwell elapsed
    _abStepDone[1] := bVacuumFb;         // 步 1 完成：真空反馈 / Step 1 done, vacuum feedback
    _abStepDone[2] := bLiftFb;           // 步 2 完成：提升到位反馈 / Step 2 done, lift feedback
    _abStepDone[3] := bOpenFb;           // 步 3 完成：开箱到位反馈 / Step 3 done, spreader feedback
    _abStepDone[4] := bFoldFb;           // 步 4 完成：折翼到位反馈 / Step 4 done, flap feedback
    _abStepDone[5] := bFoldFb;           // 步 5 完成：折后底翼共用折翼反馈 / Step 5 done, flap feedback shared
    _abStepDone[6] := bTuckFb;           // 步 6 完成：插底到位反馈 / Step 6 done, tuck feedback
    _abStepDone[7] := bPressFb;          // 步 7 完成：压底到位反馈 / Step 7 done, press feedback
    _abStepDone[8] := bEjectFb;          // 步 8 完成：推出到位反馈 / Step 8 done, eject feedback
    IF _abStepDone[3] AND (_ePhase = E_DL_CartonPhase.eOpening) THEN
        _bInfoOpen := TRUE;              // 开箱到位（信息级，关键节点） / Opening reached, info
    END_IF
END_IF

fbSeq(bStart := _bSeqStart, abStepDone := _abStepDone, auStepTimeout := _auStepTimeout,
      bHold := FALSE, bSingleStep := FALSE, bAdvance := FALSE,
      bAbort := (_bAbortStage >= 1),
      bReset := bReset AND (_ePhase = E_DL_CartonPhase.eFault)); // 步进器唯一调用点；复位仅故障相透传（步进器 bError 锁存型，v1.0.1 死锁修复；非故障相禁透传防误清） / The only sequencer call site; reset forwarded only in the fault phase, v1.0.1 deadlock fix

(*------------------------------------------------------------------------------
 * 段 6｜相位机（只做迁移与步进对账；输出在段 7 按相置位）
 *      Phase machine, transitions and step reconciliation only
 *-----------------------------------------------------------------------------*)
CASE _ePhase OF

    E_DL_CartonPhase.eIdle:                // 空闲：启动沿进就绪
        IF _bSeqStart THEN
            _ePhase := E_DL_CartonPhase.eReady; // 进就绪 / To ready
        END_IF

    E_DL_CartonPhase.eReady:               // 就绪：步进器推进到步 1 即转送箱坯
        IF fbSeq.bError THEN
            _ePhase := E_DL_CartonPhase.eFault; // 步超时，故障 / Step timeout, fault
        ELSIF (fbSeq.nCurrentStep = 1) THEN
            _ePhase := E_DL_CartonPhase.eFeeding; // 步进器已推进 / The sequencer advanced
        END_IF

    E_DL_CartonPhase.eFeeding:             // 送箱坯：步进器推进到步 3 即转开箱
        IF fbSeq.bError THEN
            _ePhase := E_DL_CartonPhase.eFault; // 步超时，故障 / Step timeout, fault
        ELSIF (fbSeq.nCurrentStep = 3) THEN
            _ePhase := E_DL_CartonPhase.eOpening; // 步进器已推进 / The sequencer advanced
        END_IF

    E_DL_CartonPhase.eOpening:             // 开箱：步进器推进到步 4 即转折底
        IF fbSeq.bError THEN
            _ePhase := E_DL_CartonPhase.eFault; // 步超时，故障 / Step timeout, fault
        ELSIF (fbSeq.nCurrentStep = 4) THEN
            _ePhase := E_DL_CartonPhase.eFolding; // 步进器已推进 / The sequencer advanced
        END_IF

    E_DL_CartonPhase.eFolding:             // 折底：步进器推进到步 7 即转封压
        IF fbSeq.bError THEN
            _ePhase := E_DL_CartonPhase.eFault; // 步超时，故障 / Step timeout, fault
        ELSIF (fbSeq.nCurrentStep = 7) THEN
            _ePhase := E_DL_CartonPhase.eSealing; // 步进器已推进 / The sequencer advanced
        END_IF

    E_DL_CartonPhase.eSealing:             // 封压：步进器推进到步 8 即转推出
        IF fbSeq.bError THEN
            _ePhase := E_DL_CartonPhase.eFault; // 步超时，故障 / Step timeout, fault
        ELSIF (fbSeq.nCurrentStep = 8) THEN
            _ePhase := E_DL_CartonPhase.eEjecting; // 步进器已推进 / The sequencer advanced
        END_IF

    E_DL_CartonPhase.eEjecting:            // 推出：步进器 bDone 即完成
        IF fbSeq.bError THEN
            _ePhase := E_DL_CartonPhase.eFault; // 步超时，故障 / Step timeout, fault
        ELSIF fbSeq.bDone THEN
            _bInfoDone := TRUE;            // 成型完成（信息级，拍 N 进入） / Erecting done, info
            _ePhase := E_DL_CartonPhase.eDone; // 本拍转出：进完成 / To done
        END_IF

    E_DL_CartonPhase.eDone:                // 完成：等启动撤销回空闲
        IF NOT bStart THEN
            _ePhase := E_DL_CartonPhase.eIdle; // 回空闲 / Back to idle
        END_IF

    E_DL_CartonPhase.eFault:               // 故障：复位沿且原因消失回空闲
        IF bReset AND (NOT _bCfgBad) AND (NOT fbSeq.bError) THEN
            _ePhase := E_DL_CartonPhase.eIdle; // 回空闲 / Back to idle
        END_IF

    ELSE                                   // 非法状态兜底（R21：CASE 必带 ELSE）
        _bIllegal := TRUE;                 // 标记非法状态 / Flag the illegal state
        _ePhase   := E_DL_CartonPhase.eFault; // 回故障态（段 7 全断） / Back to fault, all outputs off
END_CASE

(*------------------------------------------------------------------------------
 * 段 7｜输出置位（次序即安全：abort 拍仅真空断、缸全部撤，机检断言）
 *      Output assignment, abort scan cuts vacuum and retracts all cylinders
 *-----------------------------------------------------------------------------*)
CASE _ePhase OF
    E_DL_CartonPhase.eReady:               // 就绪：吸箱坯下降 / Ready: blank feed down
        bVacuumOn := (_bAbortStage = 0);   // 中止拍真空断 / Vacuum cut in abort
        bFeedOut  := (_bAbortStage = 0);   // 送坯输出 / Feed output
    E_DL_CartonPhase.eFeeding:             // 送箱坯：真空保持 + 提升 / Feeding: vacuum held, lift
        bVacuumOn := (_bAbortStage = 0);   // 真空保持 / Vacuum held
    E_DL_CartonPhase.eOpening:             // 开箱：撑箱缸 / Opening: spreader
        bVacuumOn := (_bAbortStage = 0);   // 真空保持 / Vacuum held
        bOpenOut  := (_bAbortStage = 0);   // 开箱输出 / Spreader output
    E_DL_CartonPhase.eFolding:             // 折底：折翼 + 插底缸 / Folding: flap and tuck
        bVacuumOn := (_bAbortStage = 0);   // 真空保持 / Vacuum held
        bFoldOut  := (_bAbortStage = 0);   // 折翼输出 / Flap output
        bTuckOut  := (_bAbortStage = 0) AND fbSeq.nCurrentStep >= 6; // 插底输出（步 6 起） / Tuck output from step 6
    E_DL_CartonPhase.eSealing:             // 封压：压底缸 / Sealing: press
        bPressOut := (_bAbortStage = 0);   // 压底输出 / Press output
    E_DL_CartonPhase.eEjecting:            // 推出：推出缸 / Ejecting: eject
        bEjectOut := (_bAbortStage = 0);   // 推出输出 / Eject output
    ELSE                                   // 其余相输出全断 / Otherwise all off
        bVacuumOn := FALSE;                // 真空断 / Vacuum off
        bFeedOut  := FALSE;                // 送坯断 / Feed off
        bOpenOut  := FALSE;                // 开箱断 / Spreader off
        bFoldOut  := FALSE;                // 折翼断 / Flap off
        bTuckOut  := FALSE;                // 插底断 / Tuck off
        bPressOut := FALSE;                // 压底断 / Press off
        bEjectOut := FALSE;                // 推出断 / Eject off
END_CASE

(*------------------------------------------------------------------------------
 * 段 8｜码位出口（故障级码 3 行内置 bError，R45/R101 配对）
 *      Code outlet, fault codes paired with bError
 *-----------------------------------------------------------------------------*)
IF _bIllegal THEN
    eErr   := 16#0005_0335;                // 故障级：状态机兜底 / Fault: state machine fallback
    bError := TRUE;                        // 置故障标志 / Raise the fault flag
ELSIF _bCfgBad THEN
    eErr   := 16#0005_0333;                // 故障级：组态非法 / Fault: illegal configuration
    bError := TRUE;                        // 置故障标志 / Raise the fault flag
ELSIF fbSeq.bError THEN
    eErr   := 16#0005_0334;                // 故障级：步超时 / Fault: step timeout
    bError := TRUE;                        // 置故障标志 / Raise the fault flag
ELSIF _bInfoDone THEN
    eErr := 16#0005_01F4;                  // 信息级：成型完成放行 / Info: erecting done
ELSIF _bInfoOpen THEN
    eErr := 16#0005_01F5;                  // 信息级：开箱到位提示 / Info: opening reached
END_IF

bValid := (NOT bError) AND (_ePhase <> E_DL_CartonPhase.eIdle); // 空闲/故障输出不可用 / Outputs unusable in idle or fault
ePhase := _ePhase;                       // 相位出口 / Phase outlet
END_FUNCTION_BLOCK
